(*
SPDX-FileCopyrightText: © 2026 Oleksandr Tiutyk <trofimich@gmail.com>
SPDX-License-Identifier: MIT
License: https://opensource.org/license/mit
*)

(*!
<summary>Verifies the testing library with an independent cyclic driver and direct expectations.</summary>
<description>
Runs sixteen scenarios in order with separate inner runners, including deliberately failed inner tests.
Keeps fixtures and the first diagnostic alive across scans. Publishes results directly to the ADS log.
Call Execute once per scan in the owning test task. AutomationRunner owns task memory cleanup.
This suite runs once per application initialization. Do not copy fixture state.
</description>
*)

{attribute 'no_assign'}
{attribute 'no_explicit_call' := 'do not call this function block directly'}
FUNCTION_BLOCK TestRunnerContractTest
VAR_STAT
	{attribute 'hide'}
	_ClassName : STRING := __POUNAME();
END_VAR
VAR CONSTANT
	//! <summary>Number of scenarios scheduled by the independent driver.</summary>
	_TestCount : DINT := 16;
	//! <summary>Maximum calls allowed for the empty runner to report completion.</summary>
	_EmptyScanLimit : UDINT := 16;
	//! <summary>Maximum calls per deadline phase on the configured 10 ms TestTask.</summary>
	_DeadlineScanLimit : UDINT := 32;
END_VAR
VAR_OUTPUT
	//! <summary>Number of completed scenarios with no outer assertion failures.</summary>
	PassedTests : DINT;
	//! <summary>Number of completed scenarios with an outer assertion failure or an unexpected exception.</summary>
	FailedTests : DINT;
	//! <summary>TRUE after every scenario has an outcome and the summary has been published.</summary>
	IsFinished : BOOL;
END_VAR
VAR
	_Scenario : TEST_RUNNER_CONTRACT_SCENARIO;
	_CaseFailed : BOOL;
	_FailureMessage : STRING(255);
END_VAR
VAR
	_Runner : MixedTestRunner;
	_Reporter : TOF_Testing.JUnitXmlReporter;
	_Configured : BOOL;
	_Calls : UDINT;
	_Repeated : BOOL;

	_FailingRun : IsolationTestRunner;
	_PassingRun : AssertionCallerTestRunner;
	_FailureReport : TOF_Testing.JUnitXmlReporter;
	_PassReport : TOF_Testing.JUnitXmlReporter;
	_IsolationConfigured : BOOL;
	_IsolationSecondRun : BOOL;
	_IsolationCalls : UDINT;

	_EmptyRun : EmptyTestRunner;
	_EmptyReport : TOF_Testing.JUnitXmlReporter;
	_EmptyConfigured : BOOL;
	_EmptyCalls : UDINT;
	_AbortRun : ReporterAbortTestRunner;
	_AbortReport : ThrowingTestReporter;
	_InvalidReport : TOF_Testing.JUnitXmlReporter;
	_AbortConfigured : BOOL;
	_AbortCalls : UDINT;
	_AbortPostCalls : UDINT;

	_DeadlineRun : DeadlineTestRunner;
	_DeadlineReport : TOF_Testing.JUnitXmlReporter;
	_DeadlineConfigured : BOOL;
	_DeadlineBusyFailureRun : BOOL;
	_DeadlineCalls : UDINT;
	_ActiveConfigurationChecked : BOOL;

	_DuplicateGroup : PairTestGroup(name := "Duplicates", parent := 0);
	_ParentGroup : SingleChildTestGroup(name := "Parent", parent := _ChildGroup);
	_ChildGroup : SingleChildTestGroup(name := "Child", parent := _ParentGroup);
	_IndexedGroup : PairTestGroup(name := "Indexed children", parent := 0);

	_AbortRecoveryReport : TOF_Testing.JUnitXmlReporter;
	_AbortRecovered : BOOL;
	_ExternalRun : ExternalRecoveryTestRunner;
	_ExternalReport : TOF_Testing.JUnitXmlReporter;
	_ExternalConfigured : BOOL;
	_ExternalRecovered : BOOL;
	_ExternalCalls : UDINT;

	_DiagnosticRun : DiagnosticTestRunner;
	_DiagnosticReport : TOF_Testing.JUnitXmlReporter;
	_DiagnosticConfigured : BOOL;
	_DiagnosticCalls : UDINT;

	_AssertionRun : AssertionTestRunner;
	_AssertionReport : TOF_Testing.JUnitXmlReporter;
	_AssertionsConfigured : BOOL;
	_AssertionCalls : UDINT;

	_XmlReport : TOF_Testing.JUnitXmlReporter;

	_RootTopologyRunner : RootTopologyTestRunner;
	_RootTopologyReport : TOF_Testing.JUnitXmlReporter;
	_RootTopologyConfigured : BOOL;
	_RootTopologyCalls : UDINT;

	_MissingConfigurationGroup : MissingChildrenTestGroup(name := "Missing configuration", parent := 0);
	_MissingConfigurationRunner : MissingChildrenTestRunner;
	_ExceptionAdsReporter : TOF_Testing.AdsLogReporter;
	_AdsSummaryReporter : CapturingAdsLogReporter;

	//! <summary>Synthetic Parent chains for path observation only; these fixtures are not executed as trees.</summary>
	_PathRoot : EmptyTestGroup(
		name := "AAAAAAAAAAAAAAAAAAAAAAAAAAAAAAAAAAAAAAAAAAAAAAAAAAAAAAAAAAAAAAAAAAAAAAAAAAAAAAAA",
		parent := 0
	);
	_PathSecond : EmptyTestGroup(
		name := "BBBBBBBBBBBBBBBBBBBBBBBBBBBBBBBBBBBBBBBBBBBBBBBBBBBBBBBBBBBBBBBBBBBBBBBBBBBBBBBB",
		parent := _PathRoot
	);
	_PathThird : EmptyTestGroup(
		name := "CCCCCCCCCCCCCCCCCCCCCCCCCCCCCCCCCCCCCCCCCCCCCCCCCCCCCCCCCCCCCCCCCCCCCCCCCCCCCCCC",
		parent := _PathSecond
	);
	_PathFourth : EmptyTestGroup(
		name := "DDDDDDDDDDDDDDDDDDDDDDDDDDDDDDDDDDDDDDDDDDDDDDDDDDDDDDDDDDDDDDDDDDDDDDDDDDDDDDDD",
		parent := _PathThird
	);
	_PathEmpty : EmptyTestGroup(name := "", parent := _PathRoot);
	_PathUnicode : TestingProbe(name := "Ω", parent := _PathEmpty);
	//! <summary>Supplies 81 characters to exercise ordinary truncation at the 80-character name input.</summary>
	_PathLongNameInput : WSTRING(81) := "AAAAAAAAAAAAAAAAAAAAAAAAAAAAAAAAAAAAAAAAAAAAAAAAAAAAAAAAAAAAAAAAAAAAAAAAAAAAAAAAB";
	_PathLongName : EmptyTestGroup(
		name := _PathLongNameInput,
		parent := 0
	);
	_ReportPathRoot : EmptyTestGroup(name := "Report root", parent := 0);
	_ReportPathMiddle : EmptyTestGroup(name := "Middle", parent := _ReportPathRoot);
	_ReportPathInner : EmptyTestGroup(name := "Inner", parent := _ReportPathMiddle);
	_PathReport : TOF_Testing.JUnitXmlReporter;
	_MetadataBoolAssertionContext : TOF_Testing.BoolAssertionContext;
	_MetadataByteAssertionContext : TOF_Testing.ByteAssertionContext;
	_MetadataDateAssertionContext : TOF_Testing.DateAssertionContext;
	_MetadataDateTimeAssertionContext : TOF_Testing.DateTimeAssertionContext;
	_MetadataDIntAssertionContext : TOF_Testing.DIntAssertionContext;
	_MetadataDWordAssertionContext : TOF_Testing.DWordAssertionContext;
	_MetadataIntAssertionContext : TOF_Testing.IntAssertionContext;
	_MetadataLIntAssertionContext : TOF_Testing.LIntAssertionContext;
	_MetadataLongDateAssertionContext : TOF_Testing.LongDateAssertionContext;
	_MetadataLongDateTimeAssertionContext : TOF_Testing.LongDateTimeAssertionContext;
	_MetadataLongRealAssertionContext : TOF_Testing.LongRealAssertionContext;
	_MetadataLongTimeAssertionContext : TOF_Testing.LongTimeAssertionContext;
	_MetadataLongTimeOfDayAssertionContext : TOF_Testing.LongTimeOfDayAssertionContext;
	_MetadataLWordAssertionContext : TOF_Testing.LWordAssertionContext;
	_MetadataPointerAssertionContext : TOF_Testing.PointerAssertionContext;
	_MetadataRealAssertionContext : TOF_Testing.RealAssertionContext;
	_MetadataSIntAssertionContext : TOF_Testing.SIntAssertionContext;
	_MetadataStringAssertionContext : TOF_Testing.StringAssertionContext;
	_MetadataTimeAssertionContext : TOF_Testing.TimeAssertionContext;
	_MetadataTimeOfDayAssertionContext : TOF_Testing.TimeOfDayAssertionContext;
	_MetadataUDIntAssertionContext : TOF_Testing.UDIntAssertionContext;
	_MetadataUIntAssertionContext : TOF_Testing.UIntAssertionContext;
	_MetadataULIntAssertionContext : TOF_Testing.ULIntAssertionContext;
	_MetadataUSIntAssertionContext : TOF_Testing.USIntAssertionContext;
	_MetadataWideStringAssertionContext : TOF_Testing.WideStringAssertionContext;
	_MetadataWordAssertionContext : TOF_Testing.WordAssertionContext;
	_OtherBoolContext : TOF_Testing.BoolAssertionContext;
END_VAR

(*!
<summary>Advances one scenario and reports its outcome after completion.</summary>
<description>
Retains the first failed expectation across pending cycles. An unexpected exception fails the active scenario.
Checks the allocation latch outside the recovery block. The caller owns task memory cleanup.
Returns immediately after all scenarios finish and publishes exactly one summary per initialization.
</description>
*)
METHOD Execute
VAR
	caseName : STRING(80);
	nextScenario : TEST_RUNNER_CONTRACT_SCENARIO;
	completed : BOOL;
	exceptionCode : __SYSTEM.ExceptionCode;
END_VAR
IF IsFinished THEN
	RETURN;
END_IF

IF _Scenario = TEST_RUNNER_CONTRACT_SCENARIO.STARTING THEN
	logResult(isError := FALSE, message := TOF_Core.Strings.Concat255('Starting ', TO_STRING(_TestCount), ' tests'));
	_Scenario := TEST_RUNNER_CONTRACT_SCENARIO.ELEMENT_TREE;

	RETURN;
END_IF

__TRY
	CASE _Scenario OF
		TEST_RUNNER_CONTRACT_SCENARIO.ELEMENT_TREE:
			caseName := 'Element tree, lifecycle, repeated run and JUnit';
			nextScenario := TEST_RUNNER_CONTRACT_SCENARIO.CASE_ISOLATION;
			completed := runAndCheck();

		TEST_RUNNER_CONTRACT_SCENARIO.CASE_ISOLATION:
			caseName := 'Each failure belongs to its receiving case';
			nextScenario := TEST_RUNNER_CONTRACT_SCENARIO.EMPTY_RUN;
			completed := checkCaseIsolation();

		TEST_RUNNER_CONTRACT_SCENARIO.EMPTY_RUN:
			caseName := 'An empty root passes with zero tests';
			nextScenario := TEST_RUNNER_CONTRACT_SCENARIO.REPORTER_ABORT;
			completed := checkEmptyRun();

		TEST_RUNNER_CONTRACT_SCENARIO.REPORTER_ABORT:
			caseName := 'A throwing reporter aborts without retry';
			nextScenario := TEST_RUNNER_CONTRACT_SCENARIO.DEADLINE;
			completed := checkReporterAbort();

		TEST_RUNNER_CONTRACT_SCENARIO.DEADLINE:
			caseName := 'A pending multi-cycle test fails at its deadline';
			nextScenario := TEST_RUNNER_CONTRACT_SCENARIO.GROUP_TOPOLOGY;
			completed := checkDeadline();

		TEST_RUNNER_CONTRACT_SCENARIO.GROUP_TOPOLOGY:
			caseName := 'Static group topology is validated before child callbacks';
			nextScenario := TEST_RUNNER_CONTRACT_SCENARIO.EXTERNAL_RECOVERY;
			completed := checkTopology();

		TEST_RUNNER_CONTRACT_SCENARIO.EXTERNAL_RECOVERY:
			caseName := 'External abort recovery can be retried for the same static tree';
			nextScenario := TEST_RUNNER_CONTRACT_SCENARIO.DIAGNOSTICS;
			completed := checkExternalRecovery();

		TEST_RUNNER_CONTRACT_SCENARIO.DIAGNOSTICS:
			caseName := 'Native and framework diagnostics outlive their exception objects';
			nextScenario := TEST_RUNNER_CONTRACT_SCENARIO.ADS_REPORTER_SUMMARY;
			completed := checkDiagnostics();

		TEST_RUNNER_CONTRACT_SCENARIO.ADS_REPORTER_SUMMARY:
			caseName := 'ADS summary retains first failure and resets on the next run';
			nextScenario := TEST_RUNNER_CONTRACT_SCENARIO.ASSERTION_CONTRACTS;
			completed := checkAdsReporterSummary();

		TEST_RUNNER_CONTRACT_SCENARIO.ASSERTION_CONTRACTS:
			caseName := 'Independent contexts, typed predicates, snapshots and chain diagnostics';
			nextScenario := TEST_RUNNER_CONTRACT_SCENARIO.XML_ENCODING;
			completed := checkAssertionContracts();

		TEST_RUNNER_CONTRACT_SCENARIO.XML_ENCODING:
			caseName := 'JUnit preserves long text and replaces forbidden Unicode sequences';
			nextScenario := TEST_RUNNER_CONTRACT_SCENARIO.RUNNER_TOPOLOGY;
			completed := checkXmlEncoding();

		TEST_RUNNER_CONTRACT_SCENARIO.RUNNER_TOPOLOGY:
			caseName := 'Static runner validates roots at startup and executes without rescanning';
			nextScenario := TEST_RUNNER_CONTRACT_SCENARIO.EXCEPTION_CLASSES;
			completed := checkRunnerTopology();

		TEST_RUNNER_CONTRACT_SCENARIO.EXCEPTION_CLASSES:
			caseName := 'Missing static storage is diagnosed before child access';
			nextScenario := TEST_RUNNER_CONTRACT_SCENARIO.CONTEXT_OBJECTS;
			completed := checkExceptionClasses();

		TEST_RUNNER_CONTRACT_SCENARIO.CONTEXT_OBJECTS:
			caseName := 'Typed contexts and concrete runner expose Object metadata and identity';
			nextScenario := TEST_RUNNER_CONTRACT_SCENARIO.PATHS;
			completed := checkContextObjects();

		TEST_RUNNER_CONTRACT_SCENARIO.PATHS:
			caseName := 'Paths follow live Parent links without Reset context';
			nextScenario := TEST_RUNNER_CONTRACT_SCENARIO.INDEXED_CHILDREN;
			completed := checkPaths();

		TEST_RUNNER_CONTRACT_SCENARIO.INDEXED_CHILDREN:
			caseName := 'Indexed children preserve order and reject missing storage or invalid indices';
			nextScenario := TEST_RUNNER_CONTRACT_SCENARIO.FINISHED;
			completed := checkIndexedChildren();
	ELSE
		caseName := 'Scenario selection';
		nextScenario := TEST_RUNNER_CONTRACT_SCENARIO.FINISHED;
		expect(condition := FALSE, message := 'Invalid scenario selection');
		completed := TRUE;
	END_CASE
__CATCH(exceptionCode)
	expect(
		condition := FALSE,
		message := TOF_Core.Strings.Concat255('Unexpected PLC exception ', TO_STRING(exceptionCode))
	);
	completed := TRUE;
__ENDTRY

TOF_Core.DynamicMemoryManager.RaiseIfAllocationFailed();

IF NOT completed THEN
	RETURN;
END_IF

IF _CaseFailed THEN
	FailedTests := FailedTests + 1;
	logResult(
		isError := TRUE,
		message := TOF_Core.Strings.Concat255(caseName, ': ', _FailureMessage)
	);
ELSE
	PassedTests := PassedTests + 1;
END_IF

_CaseFailed := FALSE;
_FailureMessage := '';
_Scenario := nextScenario;

IF _Scenario = TEST_RUNNER_CONTRACT_SCENARIO.FINISHED THEN
	logResult(
		isError := FailedTests <> 0,
		message := TOF_Core.Strings.Concat255(
			'Finished: ',
			TO_STRING(PassedTests),
			' passed, ',
			TO_STRING(FailedTests),
			' failed'
		)
	);
	IsFinished := TRUE;
END_IF
END_METHOD

(*!
<summary>Copies the first diagnostic when an expectation fails.</summary>
<param name="condition">TRUE when the expectation holds.</param>
<param name="message">Description of the failed expectation.</param>
*)
METHOD PRIVATE expect
VAR_INPUT
	condition : BOOL;
	message : STRING(255);
END_VAR
IF NOT condition AND_THEN NOT _CaseFailed THEN
	_CaseFailed := TRUE;
	_FailureMessage := message;
END_IF
END_METHOD

(*!
<summary>Checks that a predicate is false.</summary>
<param name="condition">Predicate that must be FALSE.</param>
<param name="message">Description of the failed expectation.</param>
*)
METHOD PRIVATE expectFalse
VAR_INPUT
	condition : BOOL;
	message : STRING(255);
END_VAR
expect(condition := NOT condition, message := message);
END_METHOD

(*!
<summary>Compares two DINT values and records differences.</summary>
<param name="expected">Expected value determined by the scenario.</param>
<param name="actual">Observed value.</param>
<param name="message">Description of the failed expectation.</param>
*)
METHOD PRIVATE expectDInt
VAR_INPUT
	expected : DINT;
	actual : DINT;
	message : STRING(255);
END_VAR
IF actual <> expected AND_THEN NOT _CaseFailed THEN
	expect(
		condition := FALSE,
		message := TOF_Core.Strings.Concat255(
			message,
			' (expected ',
			TO_STRING(expected),
			', actual ',
			TO_STRING(actual),
			')'
		)
	);
END_IF
END_METHOD

(*!
<summary>Compares two UDINT values and records differences.</summary>
<param name="expected">Expected value determined by the scenario.</param>
<param name="actual">Observed value.</param>
<param name="message">Description of the failed expectation.</param>
*)
METHOD PRIVATE expectUDInt
VAR_INPUT
	expected : UDINT;
	actual : UDINT;
	message : STRING(255);
END_VAR
IF actual <> expected AND_THEN NOT _CaseFailed THEN
	expect(
		condition := FALSE,
		message := TOF_Core.Strings.Concat255(
			message,
			' (expected ',
			TO_STRING(expected),
			', actual ',
			TO_STRING(actual),
			')'
		)
	);
END_IF
END_METHOD

(*!
<summary>Publishes a diagnostic without using the library under test.</summary>
<param name="isError">TRUE for scenario errors and failed summaries.</param>
<param name="message">Diagnostic to publish.</param>
*)
METHOD PRIVATE logResult
VAR_INPUT
	isError : BOOL;
	message : STRING(255);
END_VAR
VAR
	severity : DWORD;
END_VAR
severity := SEL(
	isError,
	Tc2_System.Global_Variables.ADSLOG_MSGTYPE_HINT,
	Tc2_System.Global_Variables.ADSLOG_MSGTYPE_ERROR
);

Tc2_System.ADSLOGSTR(
	msgCtrlMask := severity OR Tc2_System.Global_Variables.ADSLOG_MSGTYPE_LOG,
	msgFmtStr := '[TestRunnerContractTest] %s',
	strArg := message
);
END_METHOD

(*!
<summary>Checks a caught failure through its dedicated exception interface before task cleanup.</summary>
<description>Only borrows the exception during this call; no exception reference survives the test cycle.</description>
*)
METHOD PRIVATE assertCaughtExceptionType
VAR_INPUT
	exceptionCode : __SYSTEM.ExceptionCode;
	expectedTypeName : STRING;
END_VAR
VAR
	exception : TOF_Core.IException;
	standardException : TOF_Core.IStandardException;
	argumentNotSpecified : TOF_Core.IArgumentNotSpecifiedException;
	memberNotSpecified : TOF_Core.IDataMemberNotSpecifiedException;
	argumentValueNotSupported : TOF_Core.IArgumentValueNotSupportedException;
	argumentOutOfRange : TOF_Core.IArgumentOutOfRangeException;
	matchesType : BOOL;
END_VAR
exception := TOF_Core.ExceptionManager.GetLastException(
	exceptionCode := exceptionCode,
	catchPointNamespaceName := CurrentNamespace.Name,
	catchPointPOUName := __POUNAME(),
	catchPointPosition := __POSITION()
);
expect(condition := exception <> 0, message := 'Caught failure exposes its exception payload');

IF exception = 0 THEN
	RETURN;
END_IF

IF expectedTypeName = 'StandardException' THEN
	matchesType := __QUERYINTERFACE(exception, standardException);
ELSIF expectedTypeName = 'ArgumentNotSpecifiedException' THEN
	matchesType := __QUERYINTERFACE(exception, argumentNotSpecified);
ELSIF expectedTypeName = 'DataMemberNotSpecifiedException' THEN
	matchesType := __QUERYINTERFACE(exception, memberNotSpecified);
ELSIF expectedTypeName = 'ArgumentValueNotSupportedException' THEN
	matchesType := __QUERYINTERFACE(exception, argumentValueNotSupported);
ELSIF expectedTypeName = 'ArgumentOutOfRangeException' THEN
	matchesType := __QUERYINTERFACE(exception, argumentOutOfRange);
END_IF

expect(condition := matchesType, message := 'Exception interface matches the expected failure category');
END_METHOD

(*!
<summary>Checks concrete metadata through a borrowed Object interface.</summary>
<description>Checks namespace, class, size and address separately with distinct failure diagnostics.</description>
<param name="object">Live instance whose metadata is read without preparation.</param>
<param name="expectedNamespaceName">Namespace of the project declaring the concrete type.</param>
<param name="expectedClassName">Concrete context class name.</param>
<param name="expectedSize">Compiler-reported size of the complete concrete context.</param>
<param name="expectedAddress">Address of the concrete context, without ownership transfer.</param>
*)
METHOD PRIVATE assertObjectMetadata
VAR_INPUT
	object : TOF_Core.IObject;
	expectedNamespaceName : STRING;
	expectedClassName : STRING;
	expectedSize : ULINT;
	expectedAddress : PVOID;
END_VAR
expect(condition := object <> 0, message := expectedClassName);

IF object = 0 THEN
	RETURN;
END_IF

expect(
	condition := object.ClassName = expectedClassName,
	message := TOF_Core.Strings.Concat255(expectedClassName, ': ClassName')
);
expect(
	condition := object.NamespaceName = expectedNamespaceName,
	message := TOF_Core.Strings.Concat255(expectedClassName, ': NamespaceName')
);
expect(
	condition := object.SelfSize = expectedSize,
	message := TOF_Core.Strings.Concat255(expectedClassName, ': SelfSize')
);
expect(
	condition := object.SelfAddress = expectedAddress,
	message := TOF_Core.Strings.Concat255(expectedClassName, ': SelfAddress')
);
END_METHOD

(*!
<summary>Checks independent typed and generic contexts, native predicates and chain-wide diagnostics.</summary>
<description>Configures the persistent output probes through a local reference without copying them.
Returns TRUE when all observations for this scenario are complete.
</description>
*)
METHOD PRIVATE checkAssertionContracts : BOOL
VAR
	probe : REFERENCE TO AssertionContractProbe;
END_VAR
IF NOT _AssertionsConfigured THEN
	probe REF= _AssertionRun.Assertion0;
	probe.Scenario := ASSERTION_PROBE_SCENARIO.FLOAT_TOLERANCE;
	probe REF= _AssertionRun.Assertion1;
	probe.Scenario := ASSERTION_PROBE_SCENARIO.INTEGER_EXACT;
	probe REF= _AssertionRun.Assertion2;
	probe.Scenario := ASSERTION_PROBE_SCENARIO.TYPED_LITERALS;
	probe REF= _AssertionRun.Assertion3;
	probe.Scenario := ASSERTION_PROBE_SCENARIO.MESSAGE_CHAIN;
	probe REF= _AssertionRun.Assertion4;
	probe.Scenario := ASSERTION_PROBE_SCENARIO.NEGATIVE_TOLERANCE;
	probe REF= _AssertionRun.Assertion5;
	probe.Scenario := ASSERTION_PROBE_SCENARIO.NAN_TOLERANCE;
	probe REF= _AssertionRun.Assertion6;
	probe.Scenario := ASSERTION_PROBE_SCENARIO.INFINITE_TOLERANCE;
	probe REF= _AssertionRun.Assertion7;
	probe.Scenario := ASSERTION_PROBE_SCENARIO.MESSAGE_RESET;
	probe REF= _AssertionRun.Assertion8;
	probe.Scenario := ASSERTION_PROBE_SCENARIO.POINTERS_AND_STRINGS;
	probe REF= _AssertionRun.Assertion9;
	probe.Scenario := ASSERTION_PROBE_SCENARIO.FIRST_FAILURE;
	probe REF= _AssertionRun.Assertion10;
	probe.Scenario := ASSERTION_PROBE_SCENARIO.SPECIAL_FLOATS;
	probe REF= _AssertionRun.Assertion11;
	probe.Scenario := ASSERTION_PROBE_SCENARIO.OPPOSITE_LIMITS;
	probe REF= _AssertionRun.Assertion12;
	probe.Scenario := ASSERTION_PROBE_SCENARIO.GENERIC_MESSAGE_CHAIN;
	probe REF= _AssertionRun.Assertion13;
	probe.Scenario := ASSERTION_PROBE_SCENARIO.GENERIC_MESSAGE_RESET;
	probe REF= _AssertionRun.Assertion14;
	probe.Scenario := ASSERTION_PROBE_SCENARIO.CONTEXT_TRANSITIONS;
	probe REF= _AssertionRun.Assertion15;
	probe.Scenario := ASSERTION_PROBE_SCENARIO.TYPED_MESSAGE_AFTER_GENERIC;
	probe REF= _AssertionRun.Assertion16;
	probe.Scenario := ASSERTION_PROBE_SCENARIO.GENERIC_MESSAGE_AFTER_TYPED;
	probe REF= _AssertionRun.Assertion17;
	probe.Scenario := ASSERTION_PROBE_SCENARIO.TYPED_MESSAGE_RESET_AFTER_GENERIC;
	probe REF= _AssertionRun.Assertion18;
	probe.Scenario := ASSERTION_PROBE_SCENARIO.INTEGER_FAILURE;
	probe REF= _AssertionRun.Assertion19;
	probe.Scenario := ASSERTION_PROBE_SCENARIO.BITSTRING_FAILURE;
	probe REF= _AssertionRun.Assertion20;
	probe.Scenario := ASSERTION_PROBE_SCENARIO.POINTER_FAILURE;
	probe REF= _AssertionRun.Assertion21;
	probe.Scenario := ASSERTION_PROBE_SCENARIO.STRING_LONG_FAILURE;
	probe REF= _AssertionRun.Assertion22;
	probe.Scenario := ASSERTION_PROBE_SCENARIO.WIDE_STRING_LONG_FAILURE;
	probe REF= _AssertionRun.Assertion23;
	probe.Scenario := ASSERTION_PROBE_SCENARIO.STRING_CONTAINMENT_FAILURE;
	probe REF= _AssertionRun.Assertion24;
	probe.Scenario := ASSERTION_PROBE_SCENARIO.FLOAT_ORDERING_FAILURE;
	probe REF= _AssertionRun.Assertion25;
	probe.Scenario := ASSERTION_PROBE_SCENARIO.FLOAT_EQUALITY_FAILURE;
	probe REF= _AssertionRun.Assertion26;
	probe.Scenario := ASSERTION_PROBE_SCENARIO.TIME_ORDERING_FAILURE;
	_AssertionRun.Reporter := _AssertionReport;
	_AssertionsConfigured := TRUE;
END_IF

_AssertionRun.Execute(cleanupTaskMemory := FALSE);
_AssertionCalls := _AssertionCalls + 1;

IF NOT _AssertionRun.IsFinished AND_THEN _AssertionCalls < 32 THEN
	RETURN;
END_IF

expect(condition := _AssertionRun.IsFinished, message := 'Twenty-seven assertion leaves finish within 32 scans');
expectDInt(expected := 27, actual := _AssertionRun.TotalTests, message := 'Every assertion scenario executes');
expectDInt(
	expected := 7,
	actual := _AssertionRun.PassedTests,
	message := 'Seven supported assertion scenarios pass'
);
expectDInt(
	expected := 20,
	actual := _AssertionRun.FailedTests,
	message := 'Twenty deliberate failures are recorded'
);
expect(
	condition := _AssertionRun.Assertion0.Outcome = TOF_Testing.TEST_OUTCOME.PASSED,
	message := 'Assertion scenario 0 has its expected passed outcome'
);
expect(
	condition := _AssertionRun.Assertion1.Outcome = TOF_Testing.TEST_OUTCOME.PASSED,
	message := 'Assertion scenario 1 has its expected passed outcome'
);
expect(
	condition := _AssertionRun.Assertion2.Outcome = TOF_Testing.TEST_OUTCOME.PASSED,
	message := 'Assertion scenario 2 has its expected passed outcome'
);
expect(
	condition := _AssertionRun.Assertion3.Outcome = TOF_Testing.TEST_OUTCOME.FAILED,
	message := 'Assertion scenario 3 has its expected failed outcome'
);
expect(
	condition := _AssertionRun.Assertion4.Outcome = TOF_Testing.TEST_OUTCOME.FAILED,
	message := 'Assertion scenario 4 has its expected failed outcome'
);
expect(
	condition := _AssertionRun.Assertion5.Outcome = TOF_Testing.TEST_OUTCOME.FAILED,
	message := 'Assertion scenario 5 has its expected failed outcome'
);
expect(
	condition := _AssertionRun.Assertion6.Outcome = TOF_Testing.TEST_OUTCOME.FAILED,
	message := 'Assertion scenario 6 has its expected failed outcome'
);
expect(
	condition := _AssertionRun.Assertion7.Outcome = TOF_Testing.TEST_OUTCOME.FAILED,
	message := 'Assertion scenario 7 has its expected failed outcome'
);
expect(
	condition := _AssertionRun.Assertion8.Outcome = TOF_Testing.TEST_OUTCOME.PASSED,
	message := 'Assertion scenario 8 has its expected passed outcome'
);
expect(
	condition := _AssertionRun.Assertion9.Outcome = TOF_Testing.TEST_OUTCOME.FAILED,
	message := 'Assertion scenario 9 has its expected failed outcome'
);
expect(
	condition := _AssertionRun.Assertion10.Outcome = TOF_Testing.TEST_OUTCOME.PASSED,
	message := 'Assertion scenario 10 has its expected passed outcome'
);
expect(
	condition := _AssertionRun.Assertion11.Outcome = TOF_Testing.TEST_OUTCOME.PASSED,
	message := 'Assertion scenario 11 has its expected passed outcome'
);
expect(
	condition := _AssertionRun.Assertion12.Outcome = TOF_Testing.TEST_OUTCOME.FAILED,
	message := 'Assertion scenario 12 has its expected failed outcome'
);
expect(
	condition := _AssertionRun.Assertion13.Outcome = TOF_Testing.TEST_OUTCOME.FAILED,
	message := 'Assertion scenario 13 has its expected failed outcome'
);
expect(
	condition := _AssertionRun.Assertion9.FailureMessage = "First diagnostic",
	message := 'Later assertion and teardown exception preserve the first failure'
);
expect(
	condition := TOF_Core.WideStrings.Contains(
		stringToSearchIn := _AssertionRun.Assertion3.FailureMessage,
		stringToFind := "Chain diagnostic: Expected value < "
	),
	message := 'The message survives a successful assertion in the same typed chain'
);
expect(
	condition := NOT TOF_Core.WideStrings.Contains(
		stringToSearchIn := _AssertionRun.Assertion7.FailureMessage,
		stringToFind := "Previous diagnostic"
	),
	message := 'Omitting the typed entry message clears the previous prefix'
);
expect(
	condition := TOF_Core.WideStrings.Contains(
		stringToSearchIn := _AssertionRun.Assertion12.FailureMessage,
		stringToFind := "Generic chain diagnostic: Expected value < "
	),
	message := 'Borrowed assertions retain the same chain-wide message contract'
);
expect(
	condition := NOT TOF_Core.WideStrings.Contains(
		stringToSearchIn := _AssertionRun.Assertion13.FailureMessage,
		stringToFind := "Previous generic diagnostic"
	),
	message := 'Omitting the borrowed entry message clears the previous prefix'
);
expect(
	condition := TOF_Core.WideStrings.Contains(
		stringToSearchIn := _AssertionRun.Assertion4.FailureMessage,
		stringToFind := "finite nonnegative comparison tolerance"
	),
	message := 'An invalid tolerance fails before a comparison that would otherwise pass'
);
expect(
	condition := _AssertionRun.Assertion14.Outcome = TOF_Testing.TEST_OUTCOME.PASSED,
	message := 'Independent context scenario CONTEXT_TRANSITIONS has its expected outcome'
);
expect(
	condition := _AssertionRun.Assertion15.Outcome = TOF_Testing.TEST_OUTCOME.FAILED,
	message := 'Independent context scenario TYPED_MESSAGE_AFTER_GENERIC has its expected outcome'
);
expect(
	condition := _AssertionRun.Assertion15.FailureMessage = "Independent typed: Expected: 11, but was: 10",
	message := 'Independent context scenario TYPED_MESSAGE_AFTER_GENERIC retains its diagnostic'
);
expect(
	condition := _AssertionRun.Assertion16.Outcome = TOF_Testing.TEST_OUTCOME.FAILED,
	message := 'Independent context scenario GENERIC_MESSAGE_AFTER_TYPED has its expected outcome'
);
expect(
	condition := _AssertionRun.Assertion16.FailureMessage = "Independent generic: Expected: 2, but was: 1",
	message := 'Independent context scenario GENERIC_MESSAGE_AFTER_TYPED retains its diagnostic'
);
expect(
	condition := _AssertionRun.Assertion17.Outcome = TOF_Testing.TEST_OUTCOME.FAILED,
	message := 'Independent context scenario TYPED_MESSAGE_RESET_AFTER_GENERIC has its expected outcome'
);
expect(
	condition := _AssertionRun.Assertion17.FailureMessage = "Expected: 2, but was: 1",
	message := 'Independent context scenario TYPED_MESSAGE_RESET_AFTER_GENERIC retains its diagnostic'
);
expect(
	condition := _AssertionRun.Assertion18.Outcome = TOF_Testing.TEST_OUTCOME.FAILED,
	message := 'Independent context scenario INTEGER_FAILURE has its expected outcome'
);
expect(
	condition := _AssertionRun.Assertion18.FailureMessage = "Expected: -2, but was: -3",
	message := 'Independent context scenario INTEGER_FAILURE retains its diagnostic'
);
expect(
	condition := _AssertionRun.Assertion19.Outcome = TOF_Testing.TEST_OUTCOME.FAILED,
	message := 'Independent context scenario BITSTRING_FAILURE has its expected outcome'
);
expect(
	condition := _AssertionRun.Assertion19.FailureMessage = "Expected: 11, but was: 10",
	message := 'Independent context scenario BITSTRING_FAILURE retains its diagnostic'
);
expect(
	condition := _AssertionRun.Assertion20.Outcome = TOF_Testing.TEST_OUTCOME.FAILED,
	message := 'Independent context scenario POINTER_FAILURE has its expected outcome'
);
expect(
	condition := TOF_Core.WideStrings.Contains(
		stringToSearchIn := _AssertionRun.Assertion20.FailureMessage,
		stringToFind := "Expected: 0, but was: "
	),
	message := 'Independent context scenario POINTER_FAILURE retains its diagnostic'
);
expect(
	condition := _AssertionRun.Assertion21.Outcome = TOF_Testing.TEST_OUTCOME.FAILED,
	message := 'Independent context scenario STRING_LONG_FAILURE has its expected outcome'
);
expect(
	condition := TOF_Core.WideStrings.Contains(
		stringToSearchIn := _AssertionRun.Assertion21.FailureMessage,
		stringToFind := "ASCII expected suffix"
	),
	message := 'Independent context scenario STRING_LONG_FAILURE retains its diagnostic'
);
expect(
	condition := _AssertionRun.Assertion22.Outcome = TOF_Testing.TEST_OUTCOME.FAILED,
	message := 'Independent context scenario WIDE_STRING_LONG_FAILURE has its expected outcome'
);
expect(
	condition := TOF_Core.WideStrings.Contains(
		stringToSearchIn := _AssertionRun.Assertion22.FailureMessage,
		stringToFind := "Wide expected suffix"
	),
	message := 'Independent context scenario WIDE_STRING_LONG_FAILURE retains its diagnostic'
);
expect(
	condition := _AssertionRun.Assertion23.Outcome = TOF_Testing.TEST_OUTCOME.FAILED,
	message := 'Independent context scenario STRING_CONTAINMENT_FAILURE has its expected outcome'
);
expect(
	condition := _AssertionRun.Assertion23.FailureMessage = "Expected text to contain 'missing', but was: 'present'",
	message := 'Independent context scenario STRING_CONTAINMENT_FAILURE retains its diagnostic'
);
expect(
	condition := _AssertionRun.Assertion24.Outcome = TOF_Testing.TEST_OUTCOME.FAILED,
	message := 'Independent context scenario FLOAT_ORDERING_FAILURE has its expected outcome'
);
expect(
	condition := TOF_Core.WideStrings.Contains(
		stringToSearchIn := _AssertionRun.Assertion24.FailureMessage,
		stringToFind := "Expected value > "
	),
	message := 'Independent context scenario FLOAT_ORDERING_FAILURE retains its diagnostic'
);
expect(
	condition := _AssertionRun.Assertion25.Outcome = TOF_Testing.TEST_OUTCOME.FAILED,
	message := 'Independent context scenario FLOAT_EQUALITY_FAILURE has its expected outcome'
);
expect(
	condition := TOF_Core.WideStrings.Contains(
		stringToSearchIn := _AssertionRun.Assertion25.FailureMessage,
		stringToFind := ", tolerance: "
	),
	message := 'Independent context scenario FLOAT_EQUALITY_FAILURE retains its diagnostic'
);
expect(
	condition := _AssertionRun.Assertion26.Outcome = TOF_Testing.TEST_OUTCOME.FAILED,
	message := 'Independent context scenario TIME_ORDERING_FAILURE has its expected outcome'
);
expect(
	condition := TOF_Core.WideStrings.Contains(
		stringToSearchIn := _AssertionRun.Assertion26.FailureMessage,
		stringToFind := "Expected value >= "
	),
	message := 'Independent context scenario TIME_ORDERING_FAILURE retains its diagnostic'
);
checkAssertionContracts := TRUE;
END_METHOD

(*!
<summary>Checks assertion and direct failure routing between independent active cases.</summary>
<description>Configures the persistent output probes through local references without copying them.
Returns TRUE when all observations for this scenario are complete.
</description>
*)
METHOD PRIVATE checkCaseIsolation : BOOL
VAR
	passingProbe : REFERENCE TO AssertionIsolationProbe;
	failingProbe : REFERENCE TO AssertionIsolationProbe;
END_VAR
passingProbe REF= _PassingRun.Child;
failingProbe REF= _FailingRun.Child;

IF NOT _IsolationConfigured THEN
	passingProbe.Peer := ADR(failingProbe);
	failingProbe.Timeout := T#0S;
	passingProbe.Timeout := T#0S;
	_FailingRun.Reporter := _FailureReport;
	_PassingRun.Reporter := _PassReport;
	_IsolationConfigured := TRUE;
END_IF

_FailingRun.Execute(cleanupTaskMemory := FALSE);
_PassingRun.Execute(cleanupTaskMemory := FALSE);
_IsolationCalls := _IsolationCalls + 1;

IF NOT (_FailingRun.IsFinished AND_THEN _PassingRun.IsFinished) AND_THEN _IsolationCalls < 16 THEN
	RETURN;
END_IF

expect(condition := _FailingRun.IsFinished AND _PassingRun.IsFinished, message := 'Both runs finish');
expectDInt(expected := 1, actual := _FailingRun.FailedTests, message := 'Failure belongs to receiver');
expectDInt(expected := 1, actual := _PassingRun.PassedTests, message := 'Calling case passes');
expectDInt(expected := 0, actual := _PassingRun.FailedTests, message := 'Calling case has no peer failure');

IF NOT _IsolationSecondRun AND_THEN _FailingRun.IsFinished AND_THEN _PassingRun.IsFinished THEN
	_IsolationSecondRun := TRUE;
	passingProbe.UseDirectFailure := TRUE;
	_IsolationCalls := 0;
	_FailingRun.Reset();
	_PassingRun.Reset();
	RETURN;
END_IF

checkCaseIsolation := TRUE;
END_METHOD

(*!
<summary>Checks all typed contexts through IObject before assertion preparation.</summary>
<description>
Persistent contexts retain their default state. Checks metadata, addresses and inherited identity equality;
no test callback or Prepare call is required to read Object metadata.
Also checks concrete runner metadata, the inherited INamed signature and the constructor-copied group name.
Context namespaces are compared with an independent library reporter; runner metadata uses the consumer namespace.

Returns TRUE when all observations for this scenario are complete.
</description>
*)
METHOD PRIVATE checkContextObjects : BOOL
VAR
	first : TOF_Core.IObject;
	second : TOF_Core.IObject;
	group : TOF_Core.IObject;
	named : TOF_Core.INamed;
	displayName : REFERENCE TO WSTRING;
	concreteDisplayName : REFERENCE TO WSTRING;
END_VAR
assertObjectMetadata(
	object := _Runner,
	expectedNamespaceName := CurrentNamespace.Name,
	expectedClassName := 'MixedTestRunner',
	expectedSize := XSIZEOF(_Runner),
	expectedAddress := ADR(_Runner)
);

assertObjectMetadata(
	object := _MetadataBoolAssertionContext,
	expectedNamespaceName := _ExceptionAdsReporter.NamespaceName,
	expectedClassName := 'BoolAssertionContext',
	expectedSize := XSIZEOF(_MetadataBoolAssertionContext),
	expectedAddress := ADR(_MetadataBoolAssertionContext)
);
assertObjectMetadata(
	object := _MetadataByteAssertionContext,
	expectedNamespaceName := _ExceptionAdsReporter.NamespaceName,
	expectedClassName := 'ByteAssertionContext',
	expectedSize := XSIZEOF(_MetadataByteAssertionContext),
	expectedAddress := ADR(_MetadataByteAssertionContext)
);
assertObjectMetadata(
	object := _MetadataDateAssertionContext,
	expectedNamespaceName := _ExceptionAdsReporter.NamespaceName,
	expectedClassName := 'DateAssertionContext',
	expectedSize := XSIZEOF(_MetadataDateAssertionContext),
	expectedAddress := ADR(_MetadataDateAssertionContext)
);
assertObjectMetadata(
	object := _MetadataDateTimeAssertionContext,
	expectedNamespaceName := _ExceptionAdsReporter.NamespaceName,
	expectedClassName := 'DateTimeAssertionContext',
	expectedSize := XSIZEOF(_MetadataDateTimeAssertionContext),
	expectedAddress := ADR(_MetadataDateTimeAssertionContext)
);
assertObjectMetadata(
	object := _MetadataDIntAssertionContext,
	expectedNamespaceName := _ExceptionAdsReporter.NamespaceName,
	expectedClassName := 'DIntAssertionContext',
	expectedSize := XSIZEOF(_MetadataDIntAssertionContext),
	expectedAddress := ADR(_MetadataDIntAssertionContext)
);
assertObjectMetadata(
	object := _MetadataDWordAssertionContext,
	expectedNamespaceName := _ExceptionAdsReporter.NamespaceName,
	expectedClassName := 'DWordAssertionContext',
	expectedSize := XSIZEOF(_MetadataDWordAssertionContext),
	expectedAddress := ADR(_MetadataDWordAssertionContext)
);
assertObjectMetadata(
	object := _MetadataIntAssertionContext,
	expectedNamespaceName := _ExceptionAdsReporter.NamespaceName,
	expectedClassName := 'IntAssertionContext',
	expectedSize := XSIZEOF(_MetadataIntAssertionContext),
	expectedAddress := ADR(_MetadataIntAssertionContext)
);
assertObjectMetadata(
	object := _MetadataLIntAssertionContext,
	expectedNamespaceName := _ExceptionAdsReporter.NamespaceName,
	expectedClassName := 'LIntAssertionContext',
	expectedSize := XSIZEOF(_MetadataLIntAssertionContext),
	expectedAddress := ADR(_MetadataLIntAssertionContext)
);
assertObjectMetadata(
	object := _MetadataLongDateAssertionContext,
	expectedNamespaceName := _ExceptionAdsReporter.NamespaceName,
	expectedClassName := 'LongDateAssertionContext',
	expectedSize := XSIZEOF(_MetadataLongDateAssertionContext),
	expectedAddress := ADR(_MetadataLongDateAssertionContext)
);
assertObjectMetadata(
	object := _MetadataLongDateTimeAssertionContext,
	expectedNamespaceName := _ExceptionAdsReporter.NamespaceName,
	expectedClassName := 'LongDateTimeAssertionContext',
	expectedSize := XSIZEOF(_MetadataLongDateTimeAssertionContext),
	expectedAddress := ADR(_MetadataLongDateTimeAssertionContext)
);
assertObjectMetadata(
	object := _MetadataLongRealAssertionContext,
	expectedNamespaceName := _ExceptionAdsReporter.NamespaceName,
	expectedClassName := 'LongRealAssertionContext',
	expectedSize := XSIZEOF(_MetadataLongRealAssertionContext),
	expectedAddress := ADR(_MetadataLongRealAssertionContext)
);
assertObjectMetadata(
	object := _MetadataLongTimeAssertionContext,
	expectedNamespaceName := _ExceptionAdsReporter.NamespaceName,
	expectedClassName := 'LongTimeAssertionContext',
	expectedSize := XSIZEOF(_MetadataLongTimeAssertionContext),
	expectedAddress := ADR(_MetadataLongTimeAssertionContext)
);
assertObjectMetadata(
	object := _MetadataLongTimeOfDayAssertionContext,
	expectedNamespaceName := _ExceptionAdsReporter.NamespaceName,
	expectedClassName := 'LongTimeOfDayAssertionContext',
	expectedSize := XSIZEOF(_MetadataLongTimeOfDayAssertionContext),
	expectedAddress := ADR(_MetadataLongTimeOfDayAssertionContext)
);
assertObjectMetadata(
	object := _MetadataLWordAssertionContext,
	expectedNamespaceName := _ExceptionAdsReporter.NamespaceName,
	expectedClassName := 'LWordAssertionContext',
	expectedSize := XSIZEOF(_MetadataLWordAssertionContext),
	expectedAddress := ADR(_MetadataLWordAssertionContext)
);
assertObjectMetadata(
	object := _MetadataPointerAssertionContext,
	expectedNamespaceName := _ExceptionAdsReporter.NamespaceName,
	expectedClassName := 'PointerAssertionContext',
	expectedSize := XSIZEOF(_MetadataPointerAssertionContext),
	expectedAddress := ADR(_MetadataPointerAssertionContext)
);
assertObjectMetadata(
	object := _MetadataRealAssertionContext,
	expectedNamespaceName := _ExceptionAdsReporter.NamespaceName,
	expectedClassName := 'RealAssertionContext',
	expectedSize := XSIZEOF(_MetadataRealAssertionContext),
	expectedAddress := ADR(_MetadataRealAssertionContext)
);
assertObjectMetadata(
	object := _MetadataSIntAssertionContext,
	expectedNamespaceName := _ExceptionAdsReporter.NamespaceName,
	expectedClassName := 'SIntAssertionContext',
	expectedSize := XSIZEOF(_MetadataSIntAssertionContext),
	expectedAddress := ADR(_MetadataSIntAssertionContext)
);
assertObjectMetadata(
	object := _MetadataStringAssertionContext,
	expectedNamespaceName := _ExceptionAdsReporter.NamespaceName,
	expectedClassName := 'StringAssertionContext',
	expectedSize := XSIZEOF(_MetadataStringAssertionContext),
	expectedAddress := ADR(_MetadataStringAssertionContext)
);
assertObjectMetadata(
	object := _MetadataTimeAssertionContext,
	expectedNamespaceName := _ExceptionAdsReporter.NamespaceName,
	expectedClassName := 'TimeAssertionContext',
	expectedSize := XSIZEOF(_MetadataTimeAssertionContext),
	expectedAddress := ADR(_MetadataTimeAssertionContext)
);
assertObjectMetadata(
	object := _MetadataTimeOfDayAssertionContext,
	expectedNamespaceName := _ExceptionAdsReporter.NamespaceName,
	expectedClassName := 'TimeOfDayAssertionContext',
	expectedSize := XSIZEOF(_MetadataTimeOfDayAssertionContext),
	expectedAddress := ADR(_MetadataTimeOfDayAssertionContext)
);
assertObjectMetadata(
	object := _MetadataUDIntAssertionContext,
	expectedNamespaceName := _ExceptionAdsReporter.NamespaceName,
	expectedClassName := 'UDIntAssertionContext',
	expectedSize := XSIZEOF(_MetadataUDIntAssertionContext),
	expectedAddress := ADR(_MetadataUDIntAssertionContext)
);
assertObjectMetadata(
	object := _MetadataUIntAssertionContext,
	expectedNamespaceName := _ExceptionAdsReporter.NamespaceName,
	expectedClassName := 'UIntAssertionContext',
	expectedSize := XSIZEOF(_MetadataUIntAssertionContext),
	expectedAddress := ADR(_MetadataUIntAssertionContext)
);
assertObjectMetadata(
	object := _MetadataULIntAssertionContext,
	expectedNamespaceName := _ExceptionAdsReporter.NamespaceName,
	expectedClassName := 'ULIntAssertionContext',
	expectedSize := XSIZEOF(_MetadataULIntAssertionContext),
	expectedAddress := ADR(_MetadataULIntAssertionContext)
);
assertObjectMetadata(
	object := _MetadataUSIntAssertionContext,
	expectedNamespaceName := _ExceptionAdsReporter.NamespaceName,
	expectedClassName := 'USIntAssertionContext',
	expectedSize := XSIZEOF(_MetadataUSIntAssertionContext),
	expectedAddress := ADR(_MetadataUSIntAssertionContext)
);
assertObjectMetadata(
	object := _MetadataWideStringAssertionContext,
	expectedNamespaceName := _ExceptionAdsReporter.NamespaceName,
	expectedClassName := 'WideStringAssertionContext',
	expectedSize := XSIZEOF(_MetadataWideStringAssertionContext),
	expectedAddress := ADR(_MetadataWideStringAssertionContext)
);
assertObjectMetadata(
	object := _MetadataWordAssertionContext,
	expectedNamespaceName := _ExceptionAdsReporter.NamespaceName,
	expectedClassName := 'WordAssertionContext',
	expectedSize := XSIZEOF(_MetadataWordAssertionContext),
	expectedAddress := ADR(_MetadataWordAssertionContext)
);

first := _MetadataBoolAssertionContext;
second := _OtherBoolContext;
expect(condition := first.Equals(other := first), message := 'A context equals itself');
expectFalse(condition := first.Equals(other := second), message := 'Equal snapshots do not merge context identity');
expectFalse(condition := first.Equals(other := 0), message := 'A context is distinct from null');

group := _Runner.Empty;
expect(condition := group.ClassName <> '', message := 'A concrete group provides its class name');
expect(
	condition := group.NamespaceName = _Runner.NamespaceName,
	message := 'Group and runner share the consumer namespace'
);
expect(condition := group.SelfSize = XSIZEOF(_Runner.Empty), message := 'Group size includes its concrete storage');
expect(
	condition := group.SelfAddress = ADR(_Runner.Empty),
	message := 'Group identity points to the concrete instance'
);

named := _Runner.Empty;
displayName REF= named.Name;
concreteDisplayName REF= _Runner.Empty.Name;
expect(condition := __ISVALIDREF(displayName), message := 'INamed provides a valid name reference');
expect(condition := ADR(displayName) = ADR(concreteDisplayName), message := 'INamed borrows the same name storage');
expect(condition := displayName = "Empty", message := 'INamed exposes the constructor-copied group name');

checkContextObjects := TRUE;
END_METHOD

(*!
<summary>Checks deadline completion, BUSY failure termination and mutation guards.</summary>
<description>
Configures the persistent output leaf through a local reference without copying it.
The first run must exercise active mutation guards before the deadline. The second injects a BUSY failure.
Returns TRUE when all observations for this scenario are complete.
</description>
*)
METHOD PRIVATE checkDeadline : BOOL
VAR
	deadlineProbe : REFERENCE TO AssertionIsolationProbe;
	exceptionCode : __SYSTEM.ExceptionCode;
	rejected : BOOL;
	actualParent : TOF_Testing.ITestElement;
END_VAR
deadlineProbe REF= _DeadlineRun.DeadlineGroup.Child;

IF NOT _DeadlineConfigured THEN
	deadlineProbe.CompleteAfterCycle := 0;
	deadlineProbe.Timeout := T#1MS;
	_DeadlineRun.Reporter := _DeadlineReport;
	_DeadlineConfigured := TRUE;
END_IF

_DeadlineRun.Execute(cleanupTaskMemory := FALSE);
_DeadlineCalls := _DeadlineCalls + 1;

IF deadlineProbe.IsRunning AND_THEN NOT _DeadlineBusyFailureRun AND_THEN NOT _ActiveConfigurationChecked THEN

	__TRY
		deadlineProbe.Timeout := T#2S;
	__CATCH(exceptionCode)
		assertCaughtExceptionType(
			exceptionCode := exceptionCode,
			expectedTypeName := 'StandardException'
		);
		rejected := TRUE;
	__ENDTRY

	expect(condition := rejected, message := 'An active deadline cannot be changed');
	expect(
		condition := deadlineProbe.Timeout = T#1MS,
		message := 'Rejected mutation preserves the deadline'
	);
	_DeadlineRun.Reset();
	expect(
		condition := deadlineProbe.IsRunning AND_THEN NOT _DeadlineRun.IsFinished,
		message := 'Active Reset leaves the pending leaf running'
	);
	rejected := FALSE;

	__TRY
		_DeadlineRun.Reporter := _DeadlineReport;
	__CATCH(exceptionCode)
		assertCaughtExceptionType(
			exceptionCode := exceptionCode,
			expectedTypeName := 'StandardException'
		);
		rejected := TRUE;
	__ENDTRY

	expect(condition := rejected, message := 'Active runner rejects Reporter mutation');
	actualParent := deadlineProbe.Parent;
	expect(
		condition := actualParent = _DeadlineRun.Children[0],
		message := 'The active leaf retains its constructor-assigned parent'
	);
	_ActiveConfigurationChecked := TRUE;
END_IF

IF NOT _DeadlineRun.IsFinished AND_THEN _DeadlineCalls < _DeadlineScanLimit THEN
	RETURN;
END_IF

IF NOT _DeadlineBusyFailureRun THEN
	expect(condition := _DeadlineRun.IsFinished, message := 'A one-millisecond nominal deadline terminates');
	expect(condition := _ActiveConfigurationChecked, message := 'Deadline run exercises the active mutation guards');
	expectDInt(expected := 1, actual := _DeadlineRun.FailedTests, message := 'Deadline is one failed leaf');
	expectUDInt(
		expected := 1,
		actual := deadlineProbe.TeardownCalls,
		message := 'Deadline cleanup occurs once'
	);

	IF _DeadlineRun.IsFinished THEN
		_DeadlineBusyFailureRun := TRUE;
		_DeadlineCalls := 0;
		_DeadlineRun.Reset();
		deadlineProbe.Timeout := T#0S;
		deadlineProbe.FailSelfWhileBusy := TRUE;
		RETURN;
	END_IF
ELSE
	expect(condition := _DeadlineRun.IsFinished, message := 'A failed BUSY step terminates immediately');
	expectDInt(expected := 1, actual := _DeadlineRun.FailedTests, message := 'BUSY failure counts once');
	expectUDInt(
		expected := 1,
		actual := deadlineProbe.BodyCalls,
		message := 'Failed BUSY step does not run another body cycle'
	);
	expectUDInt(
		expected := 1,
		actual := deadlineProbe.TeardownCalls,
		message := 'Failed BUSY cleanup occurs once'
	);
END_IF

checkDeadline := TRUE;
END_METHOD

(*!
<summary>Checks copied native, fallback and long diagnostics after earlier task-cycle cleanup.</summary>
<description>
Requires the inner run to finish and publish its report before the suite accepts the diagnostic results.
Returns TRUE when all observations for this scenario are complete.
</description>
*)
METHOD PRIVATE checkDiagnostics : BOOL
VAR
	probe : REFERENCE TO DiagnosticProbe;
END_VAR
IF NOT _DiagnosticConfigured THEN
	probe REF= _DiagnosticRun.NativeDiagnostic;
	probe.ThrowNative := TRUE;
	probe REF= _DiagnosticRun.FormatterDiagnostic;
	probe.ThrowOnGetMessage := TRUE;
	_DiagnosticRun.Reporter := _DiagnosticReport;
	_DiagnosticConfigured := TRUE;
END_IF

_DiagnosticRun.Execute(cleanupTaskMemory := FALSE);
_DiagnosticCalls := _DiagnosticCalls + 1;

IF NOT _DiagnosticRun.IsFinished AND_THEN _DiagnosticCalls < 16 THEN
	RETURN;
END_IF

expect(condition := _DiagnosticRun.IsFinished, message := 'The diagnostic run finishes within 16 scans');
expect(condition := _DiagnosticReport.IsReady, message := 'The diagnostic report is complete');
expectDInt(
	expected := 3,
	actual := _DiagnosticRun.FailedTests,
	message := 'All injected errors are failed leaves'
);
expect(
	condition := TOF_Core.WideStrings.Contains(stringToSearchIn := _DiagnosticRun.NativeDiagnostic.FailureMessage,
		stringToFind := "ExecuteTest"),
	message := 'Native diagnostic has the interrupted stage'
);
expect(
	condition := TOF_Core.WideStrings.Contains(stringToSearchIn := _DiagnosticRun.FormatterDiagnostic.FailureMessage,
		stringToFind := "diagnostic unavailable"),
	message := 'Failing GetMessage retains stage/code fallback'
);
expect(
	condition := TOF_Core.WideStrings.Contains(stringToSearchIn := _DiagnosticRun.LongDiagnostic.FailureMessage,
		stringToFind := "END_OF_LONG_DIAGNOSTIC"),
	message := 'Long copied exception message is not narrowed to 255'
);
expectUDInt(
	expected := 1,
	actual := _DiagnosticRun.FormatterDiagnostic.TeardownCalls,
	message := 'Fallback still tears down once'
);
checkDiagnostics := TRUE;
END_METHOD

(*!
<summary>Checks a zero-child runner completes successfully with zero tests.</summary>
<description>Returns TRUE when all observations for this scenario are complete.</description>
*)
METHOD PRIVATE checkEmptyRun : BOOL
IF NOT _EmptyConfigured THEN
	_EmptyRun.Reporter := _EmptyReport;
	_EmptyConfigured := TRUE;
END_IF

_EmptyRun.Execute(cleanupTaskMemory := FALSE);
_EmptyCalls := _EmptyCalls + 1;

IF NOT _EmptyRun.IsFinished AND_THEN _EmptyCalls < _EmptyScanLimit THEN
	RETURN;
END_IF

expect(condition := _EmptyRun.IsFinished, message := 'An empty run must finish within the scan limit');
expect(condition := _EmptyRun.AllPassed, message := 'An empty run passes');
expectDInt(expected := 0, actual := _EmptyRun.TotalTests, message := 'No synthetic empty test');
checkEmptyRun := TRUE;
END_METHOD

(*!
<summary>Checks missing static storage, safe abort recovery rejection and invalid reporter outcomes.</summary>
<description>Returns TRUE when all observations for this scenario are complete.</description>
*)
METHOD PRIVATE checkExceptionClasses : BOOL
VAR
	exceptionCode : __SYSTEM.ExceptionCode;
	rejected : BOOL;
	diagnostic : TOF_Core.ERROR_MESSAGE;
END_VAR
__TRY
	_MissingConfigurationGroup.Reset(reporter := 0);
__CATCH(exceptionCode)
	assertCaughtExceptionType(exceptionCode := exceptionCode, expectedTypeName := 'DataMemberNotSpecifiedException');
	rejected := TRUE;
__ENDTRY

expect(condition := rejected, message := 'Group Reset rejects missing child-array storage');
_MissingConfigurationRunner.Execute(cleanupTaskMemory := FALSE);
expectDInt(
	expected := -1,
	actual := _MissingConfigurationRunner.ExitCode,
	message := 'Missing runner storage aborts'
);
assertCaughtExceptionType(
	exceptionCode := _MissingConfigurationRunner.CallbackException,
	expectedTypeName := 'DataMemberNotSpecifiedException'
);
rejected := FALSE;

__TRY
	_MissingConfigurationRunner.Reset();
__CATCH(exceptionCode)
	assertCaughtExceptionType(exceptionCode := exceptionCode, expectedTypeName := 'DataMemberNotSpecifiedException');
	rejected := TRUE;
__ENDTRY

expect(condition := rejected, message := 'Recovery rejects missing storage before any child access');
expectDInt(
	expected := -1,
	actual := _MissingConfigurationRunner.ExitCode,
	message := 'Invalid recovery retains abort'
);
rejected := FALSE;

__TRY
	_ExceptionAdsReporter.ReportTestCaseResult(
		groupPath := "",
		testName := "Invalid ADS outcome",
		outcome := TOF_Testing.TEST_OUTCOME.RUNNING,
		duration := T#0S,
		message := diagnostic
	);
__CATCH(exceptionCode)
	assertCaughtExceptionType(exceptionCode := exceptionCode, expectedTypeName := 'ArgumentValueNotSupportedException');
	rejected := TRUE;
__ENDTRY

expect(condition := rejected, message := 'Reporter rejects the actual nonterminal enum value');
checkExceptionClasses := TRUE;
END_METHOD

(*!
<summary>Verifies first-failure summary retention and per-run reset through the ADS reporter callbacks.</summary>
<description>Checks rejected writes, bounded ADS output for a root leaf, and reset on the next run.
Returns TRUE when all observations for this scenario are complete.
</description>
*)
METHOD PRIVATE checkAdsReporterSummary : BOOL
VAR
	diagnostic : TOF_Core.ERROR_MESSAGE;
END_VAR
_AdsSummaryReporter.ReportRunStart(testCount := 2);
_AdsSummaryReporter.RejectWrites := TRUE;
diagnostic := "Synthetic first diagnostic";
_AdsSummaryReporter.ReportTestCaseResult(
	groupPath := "Reporter regression",
	testName := "First leaf",
	outcome := TOF_Testing.TEST_OUTCOME.FAILED,
	duration := T#0S,
	message := diagnostic
);

_AdsSummaryReporter.RejectWrites := FALSE;
diagnostic := "Synthetic second diagnostic";
_AdsSummaryReporter.ReportTestCaseResult(
	groupPath := "Reporter regression",
	testName := "Second leaf",
	outcome := TOF_Testing.TEST_OUTCOME.FAILED,
	duration := T#0S,
	message := diagnostic
);

_AdsSummaryReporter.ReportRunEnd(
	totalTests := 2,
	passedTests := 0,
	failedTests := 2,
	skippedTests := 0,
	duration := T#0S
);

expect(
	condition := _AdsSummaryReporter.LastRunSummary =
		"[TOF_Testing] Finished: 0 passed, 2 failed, 0 skipped | First failure: First leaf: Synthetic first diagnostic",
	message := 'A second failure must preserve the first failure in the summary'
);

expect(
	condition := _AdsSummaryReporter.AcceptedMessage =
		"[TOF_Testing] Finished: 0 passed, 2 failed, 0 skipped | First failed test: First leaf",
	message := 'The completion record must identify the first failure even after its detail write is rejected'
);
expect(
	condition := _AdsSummaryReporter.FailedLogWriteCount = 1,
	message := 'Exactly one rejected write must be counted'
);
expect(
	condition := _AdsSummaryReporter.LastLogFailureMessage =
		"[TOF_Testing] Reporter regression/First leaf: Synthetic first diagnostic",
	message := 'Later accepted writes must preserve the rejected message'
);

_AdsSummaryReporter.ReportRunStart(testCount := 0);

expect(
	condition := _AdsSummaryReporter.LastRunSummary = "",
	message := 'Starting a new run must clear the retained summary'
);
expect(
	condition := _AdsSummaryReporter.FailedLogWriteCount = 0 AND_THEN _AdsSummaryReporter.LastLogFailureMessage = "",
	message := 'A successful start must clear earlier failed-write observations'
);

_AdsSummaryReporter.ReportRunEnd(
	totalTests := 0,
	passedTests := 0,
	failedTests := 0,
	skippedTests := 0,
	duration := T#0S
);

expect(
	condition := _AdsSummaryReporter.LastRunSummary = "[TOF_Testing] Finished: 0 passed, 0 failed, 0 skipped",
	message := 'An empty run must omit the earlier failure'
);

_AdsSummaryReporter.ReportRunStart(testCount := 1);
diagnostic := "Long diagnostic containing a literal %s. ";
TOF_Core.WideStrings.AppendFit255(
	diagnostic,
	"AAAAAAAAAAAAAAAAAAAAAAAAAAAAAAAAAAAAAAAAAAAAAAAAAAAAAAAAAAAAAAAAAAAAAAAAAAAAAAAA",
	"BBBBBBBBBBBBBBBBBBBBBBBBBBBBBBBBBBBBBBBBBBBBBBBBBBBBBBBBBBBBBBBBBBBBBBBBBBBBBBBB",
	"CCCCCCCCCCCCCCCCCCCCCCCCCCCCCCCCCCCCCCCCCCCCCCCCCCCCCCCCCCCCCCCCCCCCCCCCCCCCCCCC"
);
_AdsSummaryReporter.ReportTestCaseResult(
	groupPath := "",
	testName := "Long failure",
	outcome := TOF_Testing.TEST_OUTCOME.FAILED,
	duration := T#0S,
	message := diagnostic
);

expect(
	condition := TOF_Core.WideStrings.GetLength(value := _AdsSummaryReporter.AcceptedMessage) = 200,
	message := 'A long ADS diagnostic must fit within the reporter limit'
);
expect(
	condition := Tc2_Standard.WLEFT(STR := _AdsSummaryReporter.AcceptedMessage, SIZE := 27) =
		"[TOF_Testing] Long failure:",
	message := 'A root leaf is logged without a leading group separator'
);

_AdsSummaryReporter.RejectWrites := TRUE;
_AdsSummaryReporter.ReportRunEnd(
	totalTests := 1,
	passedTests := 0,
	failedTests := 1,
	skippedTests := 0,
	duration := T#0S
);
expect(
	condition := _AdsSummaryReporter.LastLogFailureMessage =
		"[TOF_Testing] Finished: 0 passed, 1 failed, 0 skipped | First failed test: Long failure",
	message := 'Rejection must retain the exact completion record independently of diagnostic length'
);
expect(
	condition := _AdsSummaryReporter.FailedLogWriteCount = 1,
	message := 'A rejected completion record must be counted once'
);
_AdsSummaryReporter.RejectWrites := FALSE;

checkAdsReporterSummary := TRUE;
END_METHOD

(*!
<summary>Recovers a throwing external child, including a failed first recovery attempt.</summary>
<description>Explicitly releases the modeled resource before requesting reset recovery.
Returns TRUE when all observations for this scenario are complete.
</description>
*)
METHOD PRIVATE checkExternalRecovery : BOOL
VAR
	exceptionCode : __SYSTEM.ExceptionCode;
	rejected : BOOL;
	externalCase : REFERENCE TO ExternalElementProbe;
	actualParent : TOF_Testing.ITestElement;
END_VAR
IF NOT _ExternalConfigured THEN
	_ExternalRun.Reporter := _ExternalReport;
	_ExternalConfigured := TRUE;
END_IF

_ExternalRun.Execute(cleanupTaskMemory := FALSE);
_ExternalCalls := _ExternalCalls + 1;

IF NOT _ExternalRun.IsFinished THEN
	IF _ExternalCalls < 16 THEN
		RETURN;
	END_IF

	expect(condition := FALSE, message := 'The external recovery run must finish within 16 scans');
	_ExternalRun.ExternalCase.ReleaseResource();
	checkExternalRecovery := TRUE;

	RETURN;
END_IF

IF NOT _ExternalRecovered THEN
	expectDInt(expected := -1, actual := _ExternalRun.ExitCode, message := 'External child aborts');
	expect(
		condition := _ExternalRun.ExternalCase.ResourceActive,
		message := 'Abort does not silently release user resources'
	);
	_ExternalRun.Execute(cleanupTaskMemory := FALSE);
	expectUDInt(
		expected := 1,
		actual := _ExternalRun.ExternalCase.ExecuteCalls,
		message := 'The aborted callback is not retried before explicit recovery'
	);
	externalCase REF= _ExternalRun.ExternalCase;
	externalCase.ReleaseResource();
	expectFalse(
		condition := externalCase.ResourceActive,
		message := 'Explicit resource release completes before reset recovery'
	);
	externalCase.ThrowOnReset := TRUE;

	__TRY
		_ExternalRun.Reset();
	__CATCH(exceptionCode)
		assertCaughtExceptionType(
			exceptionCode := exceptionCode,
			expectedTypeName := 'StandardException'
		);
		rejected := TRUE;
	__ENDTRY

	expect(condition := rejected, message := 'Custom recovery Reset failure propagates');
	expectDInt(expected := -1, actual := _ExternalRun.ExitCode, message := 'Failed recovery retains abort');
	externalCase.ThrowOnReset := FALSE;
	externalCase.ThrowOnExecute := FALSE;
	_ExternalRun.Reset();
	actualParent := _ExternalRun.ExternalCase.Parent;
	expect(condition := actualParent = 0, message := 'The recovered root remains parentless');
	expectUDInt(
		expected := 3,
		actual := _ExternalRun.ExternalCase.ResetCalls,
		message := 'Failed reset was retried'
	);
	_ExternalRecovered := TRUE;
	_ExternalCalls := 0;
	RETURN;
END_IF

expect(condition := _ExternalRun.AllPassed, message := 'The same static tree succeeds after explicit recovery');
expectDInt(expected := 1, actual := _ExternalRun.PassedTests, message := 'The recovered root contributes one leaf');
expect(condition := _ExternalReport.IsReady, message := 'The recovered run completes its report');
expectUDInt(
	expected := 2,
	actual := _ExternalRun.ExternalCase.ExecuteCalls,
	message := 'Execute resumes only in the new run'
);
checkExternalRecovery := TRUE;
END_METHOD

(*!
<summary>Checks direct-child interface dispatch, fixed ordering and explicit accessor failures.</summary>
<description>
Borrows persistent fixtures before execution and after a rejected Reset. Test-only slot corruption is restored
before returning. Child identity is compared through ITestElement on both sides; indexed observation
invokes no child body.

Returns TRUE when all observations for this scenario are complete.
</description>
*)
METHOD PRIVATE checkIndexedChildren : BOOL
VAR
	element : TOF_Testing.ITestElement;
	parentElement : TOF_Testing.IParentTestElement;
	child : TOF_Testing.ITestElement;
	expectedChild : TOF_Testing.ITestElement;
	supportsChildren : BOOL;
	exceptionCode : __SYSTEM.ExceptionCode;
	rejected : BOOL;
	firstBodyCalls : UDINT;
END_VAR
element := _IndexedGroup;
supportsChildren := __QUERYINTERFACE(element, parentElement);
expect(condition := supportsChildren, message := 'A group exposes the direct-child capability');

IF NOT supportsChildren THEN
	checkIndexedChildren := TRUE;
	RETURN;
END_IF

firstBodyCalls := _IndexedGroup.First.BodyCalls;
expect(condition := parentElement.ChildCount = 2, message := 'The capability reports the fixed direct count');
expectedChild := _IndexedGroup.First;
child := parentElement.GetChildByIndex(index := 0);
expect(condition := child = expectedChild, message := 'Index zero borrows the first child');
expectedChild := _IndexedGroup.Second;
child := parentElement.GetChildByIndex(index := 1);
expect(condition := child = expectedChild, message := 'The last valid index borrows the last child');

__TRY
	child := parentElement.GetChildByIndex(index := 2);
__CATCH(exceptionCode)
	assertCaughtExceptionType(exceptionCode := exceptionCode, expectedTypeName := 'ArgumentOutOfRangeException');
	rejected := TRUE;
__ENDTRY

expect(condition := rejected, message := 'Index equal to ChildCount is rejected');
rejected := FALSE;

__TRY
	child := parentElement.GetChildByIndex(index := TOF_Core.SignedInt16.MAX_VALUE);
__CATCH(exceptionCode)
	assertCaughtExceptionType(exceptionCode := exceptionCode, expectedTypeName := 'ArgumentOutOfRangeException');
	rejected := TRUE;
__ENDTRY

expect(condition := rejected, message := 'The largest representable index is rejected before indexing');
parentElement := _Runner.Empty;
expect(condition := parentElement.ChildCount = TOF_Core.SignedInt16.ZERO, message := 'An empty group reports zero direct children');
rejected := FALSE;

__TRY
	child := parentElement.GetChildByIndex(index := 0);
__CATCH(exceptionCode)
	assertCaughtExceptionType(exceptionCode := exceptionCode, expectedTypeName := 'ArgumentOutOfRangeException');
	rejected := TRUE;
__ENDTRY

expect(condition := rejected, message := 'A valid empty array has no valid child index');
parentElement := _MissingConfigurationGroup;
rejected := FALSE;

__TRY
	child := parentElement.GetChildByIndex(index := TOF_Core.SignedInt16.MAX_VALUE);
__CATCH(exceptionCode)
	assertCaughtExceptionType(exceptionCode := exceptionCode, expectedTypeName := 'DataMemberNotSpecifiedException');
	rejected := TRUE;
__ENDTRY

expect(condition := rejected, message := 'Missing storage is diagnosed before an invalid index');

// A failed Reset does not prevent observing an existing slot; the missing selected slot remains an error.
_IndexedGroup.Children[1] := 0;
rejected := FALSE;

__TRY
	_IndexedGroup.Reset(reporter := 0);
__CATCH(exceptionCode)
	assertCaughtExceptionType(exceptionCode := exceptionCode, expectedTypeName := 'DataMemberNotSpecifiedException');
	rejected := TRUE;
__ENDTRY

expect(condition := rejected, message := 'The injected missing slot rejects Reset');
parentElement := _IndexedGroup;
expectedChild := _IndexedGroup.First;
child := parentElement.GetChildByIndex(index := 0);
expect(condition := child = expectedChild, message := 'An existing slot can be observed after failed Reset');
rejected := FALSE;

__TRY
	child := parentElement.GetChildByIndex(index := 1);
__CATCH(exceptionCode)
	assertCaughtExceptionType(exceptionCode := exceptionCode, expectedTypeName := 'DataMemberNotSpecifiedException');
	rejected := TRUE;
__ENDTRY

expect(condition := rejected, message := 'A null selected slot is a missing member');
_IndexedGroup.Children[1] := _IndexedGroup.Second;
expectUDInt(
	expected := firstBodyCalls,
	actual := _IndexedGroup.First.BodyCalls,
	message := 'Indexed observation invokes no child body'
);
_IndexedGroup.Reset(reporter := 0);
checkIndexedChildren := TRUE;
END_METHOD

(*!
<summary>Checks live root-to-element paths independently of Reset and reporting.</summary>
<description>
Checks interface dispatch, own-name inclusion, empty names, Unicode, root-prefix truncation and cycles among ancestors.
Synthetic parent-only chains isolate GetPath; they are never registered or executed as group compositions.
The existing nested and repeated-run cases independently check JUnit group paths without the leaf name.

Returns TRUE when all observations for this scenario are complete.
</description>
*)
METHOD PRIVATE checkPaths : BOOL
VAR
	element : TOF_Testing.ITestElement;
	named : TOF_Core.INamed;
	actualPath : WSTRING(255);
	expectedPath : WSTRING(255);
	exceptionCode : __SYSTEM.ExceptionCode;
	rejected : BOOL;
	diagnostic : TOF_Core.ERROR_MESSAGE;
	content : POINTER TO STRING;
	longName : WSTRING(81);
	expectedXmlName : STRING(255);
END_VAR
expectedPath := "AAAAAAAAAAAAAAAAAAAAAAAAAAAAAAAAAAAAAAAAAAAAAAAAAAAAAAAAAAAAAAAAAAAAAAAAAAAAAAAA";
named := _PathLongName;
expect(condition := named.Name = expectedPath, message := 'INamed retains the first 80 name characters');
actualPath := _PathLongName.GetPath();
expect(condition := actualPath = expectedPath, message := 'A root path observes the same bounded name');
longName := "AAAAAAAAAAAAAAAAAAAAAAAAAAAAAAAAAAAAAAAAAAAAAAAAAAAAAAAAAAAAAAAAAAAAAAAAAAAAAAAAB";
_PathReport.ReportRunStart(testCount := 1);
_PathReport.ReportTestCaseResult(
	groupPath := "",
	testName := longName,
	outcome := TOF_Testing.TEST_OUTCOME.PASSED,
	duration := T#0S,
	message := diagnostic
);
_PathReport.ReportRunEnd(totalTests := 1, passedTests := 1, failedTests := 0, skippedTests := 0, duration := T#0S);
content := _PathReport.ContentAddress;
expectedXmlName := TOF_Core.Strings.Concat255('name="', TO_STRING(expectedPath), '"');
expect(condition := _PathReport.IsReady AND_THEN content <> 0, message := 'The bounded-name report completes');

IF content <> 0 THEN
	expect(
		condition := TOF_Core.Strings.Contains(stringToSearchIn := content^, stringToFind := expectedXmlName),
		message := 'Reporter input retains exactly the first 80 name characters'
	);
END_IF

element := _DuplicateGroup;
actualPath := element.GetPath();
expect(condition := actualPath = "Duplicates", message := 'A root path contains its own name');
actualPath := _DuplicateGroup.First.GetPath();
expect(condition := actualPath = "Duplicates/First", message := 'A child path includes its group and own name');
actualPath := _Runner.FailureOuter.Failures.BodyFailure.GetPath();
expect(
	condition := actualPath = "Nested/Failures/Body failure",
	message := 'Ancestor names are ordered from the root'
);
actualPath := _Runner.Pass.GetPath();
expect(condition := actualPath = "", message := 'A nameless root has an empty path');
actualPath := _PathEmpty.GetPath();
expectedPath := "AAAAAAAAAAAAAAAAAAAAAAAAAAAAAAAAAAAAAAAAAAAAAAAAAAAAAAAAAAAAAAAAAAAAAAAAAAAAAAAA";
expect(condition := actualPath = expectedPath, message := 'An empty own name adds no separator');
actualPath := _PathUnicode.GetPath();
expectedPath := "AAAAAAAAAAAAAAAAAAAAAAAAAAAAAAAAAAAAAAAAAAAAAAAAAAAAAAAAAAAAAAAAAAAAAAAAAAAAAAAA/Ω";
expect(condition := actualPath = expectedPath, message := 'Empty ancestors are skipped and Unicode is preserved');
actualPath := _PathFourth.GetPath();
expectedPath := Tc2_Utilities.WCONCAT(
	STR1 := "AAAAAAAAAAAAAAAAAAAAAAAAAAAAAAAAAAAAAAAAAAAAAAAAAAAAAAAAAAAAAAAAAAAAAAAAAAAAAAAA/",
	STR2 := "BBBBBBBBBBBBBBBBBBBBBBBBBBBBBBBBBBBBBBBBBBBBBBBBBBBBBBBBBBBBBBBBBBBBBBBBBBBBBBBB/"
);
expectedPath := Tc2_Utilities.WCONCAT(
	STR1 := expectedPath,
	STR2 := "CCCCCCCCCCCCCCCCCCCCCCCCCCCCCCCCCCCCCCCCCCCCCCCCCCCCCCCCCCCCCCCCCCCCCCCCCCCCCCCC/DDDDDDDDDDD…"
);
expect(condition := actualPath = expectedPath, message := 'Overflow retains the root prefix and final ellipsis');

__TRY
	actualPath := _ParentGroup.Child.GetPath();
__CATCH(exceptionCode)
	assertCaughtExceptionType(exceptionCode := exceptionCode, expectedTypeName := 'StandardException');
	rejected := TRUE;
__ENDTRY

expect(condition := rejected, message := 'A cycle among ancestors is rejected without endless traversal');
actualPath := _ReportPathInner.GetPath();
_PathReport.ReportRunStart(testCount := 1);
_PathReport.ReportTestCaseResult(
	groupPath := actualPath,
	testName := "Leaf",
	outcome := TOF_Testing.TEST_OUTCOME.PASSED,
	duration := T#0S,
	message := diagnostic
);
_PathReport.ReportRunEnd(totalTests := 1, passedTests := 1, failedTests := 0, skippedTests := 0, duration := T#0S);
content := _PathReport.ContentAddress;
expect(condition := _PathReport.IsReady AND_THEN content <> 0, message := 'The deep-path report completes');

IF content <> 0 THEN
	expect(
		condition := TOF_Core.Strings.Contains(
			stringToSearchIn := content^,
			stringToFind := 'name="Leaf" classname="Report root/Middle/Inner"'
		),
		message := 'JUnit preserves all three group ancestors and keeps the leaf name separate'
	);
END_IF

checkPaths := TRUE;
END_METHOD

(*!
<summary>Verifies that a reporter failure aborts once after teardown and clears the reporter reference.</summary>
<description>The same leaf runs with a replacement reporter after a completed abort and Reset.
An incomplete run fails when it reaches the scan limit. Returns TRUE when the scenario has an outcome.
</description>
*)
METHOD PRIVATE checkReporterAbort : BOOL
VAR
	exceptionCode : __SYSTEM.ExceptionCode;
	rejected : BOOL;
	diagnostic : TOF_Core.ERROR_MESSAGE;
	actualParent : TOF_Testing.ITestElement;
END_VAR
IF _AbortRecovered THEN
	_AbortRun.Execute(cleanupTaskMemory := FALSE);
	_AbortCalls := _AbortCalls + 1;

	IF NOT _AbortRun.IsFinished AND_THEN _AbortCalls < 16 THEN
		RETURN;
	END_IF

	expect(condition := _AbortRun.IsFinished, message := 'The recovered reporter run finishes within 16 scans');
	expect(condition := _AbortRun.IsFinished AND_THEN _AbortRun.AllPassed,
		message := 'The same static tree passes after reporter abort');
	expectUDInt(
		expected := 1,
		actual := _AbortRun.AbortCase.BodyCalls,
		message := 'The same root executes once in the new run'
	);
	expectUDInt(expected := 1, actual := _AbortReport.ResultCalls, message := 'Old reporter is not retried');
	checkReporterAbort := TRUE;
	RETURN;
END_IF

IF NOT _AbortConfigured THEN

	__TRY
		_InvalidReport.ReportTestCaseResult(
			groupPath := "",
			testName := "Invalid outcome",
			outcome := TOF_Testing.TEST_OUTCOME.NOT_RUN,
			duration := T#0S,
			message := diagnostic
		);
	__CATCH(exceptionCode)
		assertCaughtExceptionType(
			exceptionCode := exceptionCode,
			expectedTypeName := 'ArgumentValueNotSupportedException'
		);
		rejected := TRUE;
	__ENDTRY

	expect(condition := rejected, message := 'A reporter rejects a nonterminal outcome');
	_AbortRun.Reporter := _AbortReport;
	_AbortConfigured := TRUE;
END_IF

_AbortRun.Execute(cleanupTaskMemory := FALSE);
_AbortCalls := _AbortCalls + 1;

IF NOT _AbortRun.IsFinished THEN
	IF _AbortCalls < 16 THEN
		RETURN;
	END_IF

	expect(condition := FALSE, message := 'Callback abort must terminate within 16 scans');
	checkReporterAbort := TRUE;

	RETURN;
END_IF

IF _AbortPostCalls < 2 THEN
	_AbortPostCalls := _AbortPostCalls + 1;
	RETURN;
END_IF

expectDInt(expected := -1, actual := _AbortRun.ExitCode, message := 'Callback abort has a distinct exit code');
expectUDInt(expected := 1, actual := _AbortReport.ResultCalls, message := 'The callback is never retried');
expectUDInt(
	expected := 1,
	actual := _AbortRun.AbortCase.TeardownCalls,
	message := 'Cleanup precedes result reporting'
);
expect(
	condition := _AbortRun.AbortCase.IsFinished AND_THEN _AbortRun.AbortCase.Reporter = 0,
	message := 'A completed leaf clears its reporter reference even when result delivery throws'
);
expectFalse(condition := _AbortReport.IsReady, message := 'An aborted report remains incomplete');
expect(
	condition := TOF_Core.WideStrings.Contains(stringToSearchIn := _AbortRun.CallbackMessage,
		stringToFind := "Reporter failed"),
	message := 'External callback diagnostic is copied'
);
_AbortRun.Reset();
expect(condition := _AbortRun.CallbackMessage = "", message := 'Reset clears copied callback diagnostic');
actualParent := _AbortRun.AbortCase.Parent;
expect(condition := actualParent = 0, message := 'The same root remains parentless after recovery');
_AbortRun.Reporter := _AbortRecoveryReport;
_AbortRecovered := TRUE;
_AbortCalls := 0;
END_METHOD

(*!
<summary>Checks static root validation, recovery guards and absence of cyclic topology scans.</summary>
<description>Deliberately corrupts test-only slots, restoring them before valid recovery and before execution reaches them.
Returns TRUE when all observations for this scenario are complete.
</description>
*)
METHOD PRIVATE checkRunnerTopology : BOOL
VAR
	exceptionCode : __SYSTEM.ExceptionCode;
	rejected : BOOL;
	runningRoot : REFERENCE TO AssertionIsolationProbe;
	actualParent : TOF_Testing.ITestElement;
END_VAR
IF NOT _RootTopologyConfigured THEN
	_RootTopologyRunner.Reporter := _RootTopologyReport;
	_RootTopologyRunner.RootTopologyFirst.Reset(reporter := 0);
	_RootTopologyRunner.RootTopologyFirst.Execute();
	_RootTopologyRunner.Children[1] := 0;
	_RootTopologyRunner.Execute(cleanupTaskMemory := FALSE);
	expectDInt(expected := -1, actual := _RootTopologyRunner.ExitCode, message := 'A null root aborts startup');
	assertCaughtExceptionType(
		exceptionCode := _RootTopologyRunner.CallbackException,
		expectedTypeName := 'DataMemberNotSpecifiedException'
	);
	expect(
		condition := _RootTopologyRunner.RootTopologyFirst.IsFinished,
		message := 'All direct roots are validated before the first Reset'
	);
	expectFalse(condition := _RootTopologyReport.IsReady, message := 'Invalid startup produces no completed report');
	expect(
		condition := _RootTopologyReport.ContentLength = TOF_Core.UnsignedInt32.ZERO,
		message := 'Invalid startup does not call ReportRunStart'
	);
	rejected := FALSE;

	__TRY
		_RootTopologyRunner.Reset();
	__CATCH(exceptionCode)
		assertCaughtExceptionType(exceptionCode := exceptionCode, expectedTypeName := 'DataMemberNotSpecifiedException');
		rejected := TRUE;
	__ENDTRY

	expect(condition := rejected, message := 'Recovery validates slots before dereferencing an invalid tree');
	expectDInt(
		expected := -1,
		actual := _RootTopologyRunner.ExitCode,
		message := 'Failed recovery retains abort'
	);
	_RootTopologyRunner.Children[1] := _RootTopologyRunner.RootTopologyGroup;
	_RootTopologyRunner.Reset();
	_RootTopologyRunner.Children[1] := _RootTopologyRunner.RootTopologyFirst;
	_RootTopologyRunner.Execute(cleanupTaskMemory := FALSE);
	expectDInt(
		expected := -1,
		actual := _RootTopologyRunner.ExitCode,
		message := 'Duplicate roots abort startup'
	);
	assertCaughtExceptionType(exceptionCode := _RootTopologyRunner.CallbackException, expectedTypeName := 'StandardException');
	_RootTopologyRunner.Children[1] := _RootTopologyRunner.RootTopologyGroup;
	_RootTopologyRunner.Reset();
	_RootTopologyRunner.Children[0] := _RootTopologyRunner.RootTopologyGroup.Child;
	_RootTopologyRunner.Execute(cleanupTaskMemory := FALSE);
	expectDInt(
		expected := -1,
		actual := _RootTopologyRunner.ExitCode,
		message := 'A group-owned root aborts startup'
	);
	assertCaughtExceptionType(exceptionCode := _RootTopologyRunner.CallbackException, expectedTypeName := 'StandardException');
	_RootTopologyRunner.Children[0] := _RootTopologyRunner.RootTopologyFirst;
	_RootTopologyRunner.Reset();
	_RootTopologyRunner.RootTopologyFirst.Execute();
	_RootTopologyRunner.Children[1] := _Runner.FailureOuter.Failures;
	_RootTopologyRunner.Execute(cleanupTaskMemory := FALSE);
	expectDInt(
		expected := -1,
		actual := _RootTopologyRunner.ExitCode,
		message := 'A nested group cannot also occupy a root slot'
	);
	assertCaughtExceptionType(exceptionCode := _RootTopologyRunner.CallbackException, expectedTypeName := 'StandardException');
	expect(
		condition := _RootTopologyRunner.RootTopologyFirst.IsFinished,
		message := 'Owned-group rejection occurs before the first direct Reset'
	);
	expect(
		condition := _RootTopologyReport.ContentLength = TOF_Core.UnsignedInt32.ZERO,
		message := 'Owned-group rejection does not start reporting'
	);
	rejected := FALSE;

	__TRY
		_RootTopologyRunner.Reset();
	__CATCH(exceptionCode)
		assertCaughtExceptionType(exceptionCode := exceptionCode, expectedTypeName := 'StandardException');
		rejected := TRUE;
	__ENDTRY

	expect(condition := rejected, message := 'Abort recovery also rejects a group-owned root');
	expectDInt(expected := -1, actual := _RootTopologyRunner.ExitCode, message := 'Invalid recovery retains abort');
	_RootTopologyRunner.Children[1] := _RootTopologyRunner.RootTopologyGroup;
	_RootTopologyRunner.Reset();
	runningRoot REF= _RootTopologyRunner.RunningRoot;
	runningRoot.Timeout := T#0S;
	_RootTopologyRunner.RunningRoot.Reset(reporter := 0);
	_RootTopologyRunner.RunningRoot.Execute();
	expect(condition := _RootTopologyRunner.RunningRoot.IsRunning, message := 'The active-root fixture is pending');
	_RootTopologyRunner.Children[0] := _RootTopologyRunner.RunningRoot;
	_RootTopologyRunner.Execute(cleanupTaskMemory := FALSE);
	expectDInt(
		expected := -1,
		actual := _RootTopologyRunner.ExitCode,
		message := 'An active root aborts startup'
	);
	assertCaughtExceptionType(exceptionCode := _RootTopologyRunner.CallbackException, expectedTypeName := 'StandardException');
	_RootTopologyRunner.RunningRoot.Reset(reporter := 0);
	_RootTopologyRunner.Children[0] := _RootTopologyRunner.RootTopologyFirst;
	_RootTopologyRunner.Reset();
	_RootTopologyRunner.Execute(cleanupTaskMemory := FALSE);
	expectFalse(condition := _RootTopologyRunner.IsFinished, message := 'Valid startup prepares the static roots');

	// Fault injection: restore the unused slot immediately after driving the first root.
	_RootTopologyRunner.Children[1] := 0;
	_RootTopologyRunner.Execute(cleanupTaskMemory := FALSE);
	_RootTopologyRunner.Children[1] := _RootTopologyRunner.RootTopologyGroup;
	expectDInt(
		expected := 0,
		actual := _RootTopologyRunner.ExitCode,
		message := 'Execution does not rescan root slots'
	);
	_RootTopologyConfigured := TRUE;
END_IF

_RootTopologyRunner.Execute(cleanupTaskMemory := FALSE);
_RootTopologyCalls := _RootTopologyCalls + 1;

IF NOT _RootTopologyRunner.IsFinished AND_THEN _RootTopologyCalls < 16 THEN
	RETURN;
END_IF

expect(condition := _RootTopologyRunner.IsFinished, message := 'The topology run finishes within 16 scans');
expect(
	condition := _RootTopologyRunner.IsFinished AND_THEN _RootTopologyRunner.AllPassed,
	message := 'The owned static roots execute successfully'
);
expectDInt(
	expected := 2,
	actual := _RootTopologyRunner.PassedTests,
	message := 'Two direct or nested leaves pass'
);
expectUDInt(
	expected := 1,
	actual := _RootTopologyRunner.RootTopologyFirst.BodyCalls,
	message := 'The first root executes once in the valid run'
);
expectUDInt(
	expected := 1,
	actual := _RootTopologyRunner.RootTopologyGroup.Child.BodyCalls,
	message := 'The nested group executes its owned leaf'
);
actualParent := _RootTopologyRunner.RootTopologyFirst.Parent;
expect(condition := actualParent = 0, message := 'Runner roots remain parentless');
actualParent := _RootTopologyRunner.RootTopologyGroup.Child.Parent;
expect(
	condition := actualParent <> 0,
	message := 'A nested leaf retains its constructor-assigned parent'
);
checkRunnerTopology := TRUE;
END_METHOD

(*!
<summary>Checks fixed parents, missing or repeated children, parent mismatch, cycles, ordered dispatch and repeat execution.</summary>
<description>
Fault injection deliberately mutates a test-only array between rejected operations and briefly during execution
to detect redundant validation. Restore every unused slot before execution reaches it.

Returns TRUE when all observations for this scenario are complete.
</description>
*)
METHOD PRIVATE checkTopology : BOOL
VAR
	exceptionCode : __SYSTEM.ExceptionCode;
	rejected : BOOL;
	expectedParent : TOF_Testing.ITestElement;
	actualParent : TOF_Testing.ITestElement;
END_VAR
expectedParent := _DuplicateGroup;
actualParent := _DuplicateGroup.First.Parent;
expect(condition := actualParent = expectedParent, message := 'Parent is assigned at construction');
actualParent := _DuplicateGroup.Parent;
expect(condition := actualParent = 0, message := 'A root is constructed without a parent');

// Deliberately corrupt the borrowed test-only array to inject topology faults.
// A later execution probe restores its unused slot before that slot is reached.
_DuplicateGroup.Children[1] := 0;

__TRY
	_DuplicateGroup.Reset(reporter := 0);
__CATCH(exceptionCode)
	assertCaughtExceptionType(exceptionCode := exceptionCode, expectedTypeName := 'DataMemberNotSpecifiedException');
	rejected := TRUE;
__ENDTRY

expect(condition := rejected, message := 'A null fixed child is rejected by Reset');
expectUDInt(
	expected := 0,
	actual := _DuplicateGroup.First.BodyCalls,
	message := 'No earlier child body executes'
);
rejected := FALSE;
_DuplicateGroup.Children[1] := _DuplicateGroup.First;

__TRY
	_DuplicateGroup.Reset(reporter := 0);
__CATCH(exceptionCode)
	assertCaughtExceptionType(exceptionCode := exceptionCode, expectedTypeName := 'StandardException');
	rejected := TRUE;
__ENDTRY

expect(condition := rejected, message := 'Duplicate fixed slots are rejected');
rejected := FALSE;
_DuplicateGroup.Children[1] := _RootTopologyRunner.RootTopologyGroup.Child;

__TRY
	_DuplicateGroup.Reset(reporter := 0);
__CATCH(exceptionCode)
	assertCaughtExceptionType(exceptionCode := exceptionCode, expectedTypeName := 'StandardException');
	rejected := TRUE;
__ENDTRY

expect(condition := rejected, message := 'A child assigned to another group is rejected');
actualParent := _DuplicateGroup.First.Parent;
expect(condition := actualParent = expectedParent, message := 'Rejection never changes Parent');
_DuplicateGroup.Children[1] := _DuplicateGroup.Second;
rejected := FALSE;

__TRY
	_ParentGroup.Reset(reporter := 0);
__CATCH(exceptionCode)
	assertCaughtExceptionType(exceptionCode := exceptionCode, expectedTypeName := 'StandardException');
	rejected := TRUE;
__ENDTRY

expect(condition := rejected, message := 'A cycle assigned by constructors is rejected before recursion');

_DuplicateGroup.Reset(reporter := 0);
// Fault injection: an unused slot must not be rescanned in Execute; restore before that slot is reached.
_DuplicateGroup.Children[1] := 0;
_DuplicateGroup.Execute();
expectUDInt(
	expected := 1,
	actual := _DuplicateGroup.First.BodyCalls,
	message := 'The first Execute reaches the first owned child through Children'
);
expectUDInt(
	expected := 0,
	actual := _DuplicateGroup.Second.BodyCalls,
	message := 'The first Execute does not reach the second owned child'
);
_DuplicateGroup.Children[1] := _DuplicateGroup.Second;
_DuplicateGroup.Execute();
expect(condition := _DuplicateGroup.IsFinished, message := 'A valid static group finishes without Configure');
expectDInt(expected := 2, actual := _DuplicateGroup.PassedCount, message := 'Both owned leaves pass');
_DuplicateGroup.Reset(reporter := 0);
_DuplicateGroup.Execute();
_DuplicateGroup.Execute();
expectDInt(
	expected := 2,
	actual := _DuplicateGroup.PassedCount,
	message := 'Reset supports another fixed-tree run'
);
expectUDInt(
	expected := 1,
	actual := _DuplicateGroup.First.BodyCalls,
	message := 'A repeated leaf executes once'
);
actualParent := _DuplicateGroup.First.Parent;
expect(condition := actualParent = expectedParent, message := 'Repeated runs preserve Parent');
_DuplicateGroup.Children[1] := 0;
rejected := FALSE;

__TRY
	_DuplicateGroup.Reset(reporter := 0);
__CATCH(exceptionCode)
	assertCaughtExceptionType(exceptionCode := exceptionCode, expectedTypeName := 'DataMemberNotSpecifiedException');
	rejected := TRUE;
__ENDTRY

expect(condition := rejected, message := 'Invalid topology is rejected on a later Reset too');
expect(
	condition := _DuplicateGroup.First.IsFinished,
	message := 'Validation precedes the first direct child Reset'
);
_DuplicateGroup.Children[1] := _DuplicateGroup.Second;
checkTopology := TRUE;
END_METHOD

(*!
<summary>Checks long XML diagnostics, supplementary Unicode, isolated surrogates and XML controls.</summary>
<description>Returns TRUE when all observations for this scenario are complete.</description>
*)
METHOD PRIVATE checkXmlEncoding : BOOL
VAR
	diagnostic : TOF_Core.ERROR_MESSAGE;
	characters : POINTER TO WORD;
	content : POINTER TO STRING;
	i : UDINT;
END_VAR
// U+1F600 is a surrogate pair; it is followed by an isolated high surrogate, U+0001, TAB and ampersand.
characters := ADR(diagnostic);
characters[0] := 16#D83D;
characters[1] := 16#DE00;
characters[2] := 16#D800;
characters[3] := 16#0001;
characters[4] := 16#0009;
characters[5] := 16#0026;

FOR i := 6 TO 405 DO
	characters[i] := 16#0078;
END_FOR

characters[406] := TOF_Core.UnsignedInt16.MIN_VALUE;
TOF_Core.WideStrings.AppendFit(targetString := diagnostic, sourceString := "END_OF_XML_DIAGNOSTIC");
_XmlReport.ReportRunStart(testCount := 1);
_XmlReport.ReportTestCaseResult(
	groupPath := "Wide",
	testName := "",
	outcome := TOF_Testing.TEST_OUTCOME.FAILED,
	duration := T#1250MS,
	message := diagnostic
);
_XmlReport.ReportRunEnd(totalTests := 1, passedTests := 0, failedTests := 1, skippedTests := 0, duration := T#1250MS);
content := _XmlReport.ContentAddress;
expect(condition := _XmlReport.IsReady AND_THEN content <> 0, message := 'Completed Unicode XML has a buffer');

IF content <> 0 THEN
	expect(
		condition := TOF_Core.Strings.Contains(stringToSearchIn := content^,
			stringToFind := '&#128512;&#65533;&#65533;&#9;&amp;'),
		message := 'Surrogate pair, isolated surrogate, forbidden control and tab are encoded'
	);
	expect(
		condition := TOF_Core.Strings.Contains(stringToSearchIn := content^, stringToFind := 'END_OF_XML_DIAGNOSTIC'),
		message := 'Diagnostic suffix beyond 255 characters survives'
	);
	expect(
		condition := TOF_Core.Strings.Contains(stringToSearchIn := content^, stringToFind := 'time="1.250"'),
		message := 'JUnit duration uses decimal seconds'
	);
END_IF

checkXmlEncoding := TRUE;
END_METHOD

(*!
<summary>Repeats a nested run and checks configured and completed leaf counts, cleanup and escaped JUnit output.</summary>
<description>Configures owned fixtures through borrowed references without copying their state.
Returns TRUE when all observations for this scenario are complete.
</description>
*)
METHOD PRIVATE runAndCheck : BOOL
VAR
	content : POINTER TO STRING;
	probe : REFERENCE TO TestingProbe;
	multiCycleProbe : REFERENCE TO AssertionIsolationProbe;
END_VAR
IF NOT _Configured THEN
	expectDInt(expected := 5, actual := _Runner.FailureOuter.TestCount, message := 'Nested leaf count');
	expectDInt(expected := 0, actual := _Runner.Empty.TestCount, message := 'Empty group leaf count');
	expectDInt(expected := 1, actual := _Runner.Pass.TestCount, message := 'Single-cycle leaf count');
	expectDInt(expected := 1, actual := _Runner.Multi.TestCount, message := 'Multi-cycle leaf count');

	probe REF= _Runner.FailureOuter.Failures.SetupFailure;
	probe.ThrowBeforeTest := TRUE;
	probe REF= _Runner.FailureOuter.Failures.BodyFailure;
	probe.ThrowBody := TRUE;
	probe REF= _Runner.FailureOuter.Failures.TeardownFailure;
	probe.ThrowAfterTest := TRUE;
	probe REF= _Runner.FailureOuter.Failures.ComparisonFailure;
	probe.InvalidComparison := TRUE;
	probe REF= _Runner.FailureOuter.Failures.DiagnosticFailure;
	probe.DiagnosticFailure := TRUE;
	_Runner.Reporter := _Reporter;
	multiCycleProbe REF= _Runner.Multi;
	multiCycleProbe.Timeout := T#0S;
	_Configured := TRUE;
END_IF

_Runner.Execute(cleanupTaskMemory := FALSE);
_Calls := _Calls + 1;

IF NOT _Runner.IsFinished AND_THEN _Calls < 32 THEN
	RETURN;
END_IF

expect(condition := _Runner.IsFinished, message := 'The tree finishes within 32 scans');
expectDInt(expected := 2, actual := _Runner.PassedTests, message := 'Single and multi-cycle leaves pass');
expectDInt(expected := 5, actual := _Runner.FailedTests, message := 'Five distinct leaf failures');
expectDInt(expected := 7, actual := _Runner.TotalTests, message := 'Groups add no synthetic tests');
expectDInt(expected := 5, actual := _Runner.FailureOuter.TestCount, message := 'Leaf count survives a run');
expectUDInt(
	expected := 0,
	actual := _Runner.FailureOuter.Failures.SetupFailure.BodyCalls,
	message := 'Failed setup suppresses body'
);
expectUDInt(
	expected := 1,
	actual := _Runner.FailureOuter.Failures.SetupFailure.TeardownCalls,
	message := 'Failed setup still cleans up'
);
expectUDInt(
	expected := 1,
	actual := _Runner.FailureOuter.Failures.BodyFailure.TeardownCalls,
	message := 'Thrown body cleans up'
);
expectUDInt(
	expected := 1,
	actual := _Runner.FailureOuter.Failures.TeardownFailure.TeardownCalls,
	message := 'Thrown teardown is not retried'
);
expectUDInt(
	expected := 1,
	actual := _Runner.Pass.BodyCalls,
	message := 'Single-cycle body executes once per run'
);
expectUDInt(
	expected := 3,
	actual := _Runner.Multi.BodyCalls,
	message := 'Multi-cycle state survives three scans'
);
expectDInt(
	expected := 0,
	actual := _Runner.Empty.FailedCount,
	message := 'An empty group passes without tests'
);
expect(condition := _Reporter.IsReady, message := 'JUnit output is complete');
expect(
	condition := TOF_Core.WideStrings.Contains(stringToSearchIn := _Runner.FailureOuter.Failures.SetupFailure.FailureMessage,
		stringToFind := "BeforeTest: "),
	message := 'Preparation stage survives exception capture'
);
expect(
	condition := TOF_Core.WideStrings.Contains(stringToSearchIn := _Runner.FailureOuter.Failures.BodyFailure.FailureMessage,
		stringToFind := "Body failed"),
	message := 'Framework payload survives task cleanup'
);
expect(
	condition := TOF_Core.WideStrings.Contains(stringToSearchIn := _Runner.FailureOuter.Failures.BodyFailure.FailureMessage,
		stringToFind := "ExecuteTest"),
	message := 'Framework source survives task cleanup'
);
expect(
	condition := TOF_Core.WideStrings.Contains(stringToSearchIn := _Runner.FailureOuter.Failures.TeardownFailure.FailureMessage,
		stringToFind := "Teardown failed"),
	message := 'Teardown payload is copied'
);

content := _Reporter.ContentAddress;
expect(condition := content <> 0, message := 'Completed XML exposes a buffer');

IF content <> 0 THEN
	expect(
		condition := TOF_Core.Strings.Contains(
			stringToSearchIn := content^,
			stringToFind := 'Expected value &lt; '
		),
		message := 'An incompatible borrowed comparison remains an assertion failure'
	);
	expect(
		condition := TOF_Core.Strings.Contains(stringToSearchIn := content^, stringToFind := '&#1070;&amp;&lt;'),
		message := 'Cyrillic and XML markup are preserved'
	);
	expect(
		condition := TOF_Core.Strings.Contains(stringToSearchIn := content^, stringToFind := 'name=""'),
		message := 'Empty test name serializes safely'
	);
	expect(
		condition := TOF_Core.Strings.Contains(stringToSearchIn := content^, stringToFind := 'classname="Nested/Failures"'),
		message := 'The nested group path is preserved'
	);
END_IF

IF NOT _Repeated AND_THEN _Runner.IsFinished THEN
	_Repeated := TRUE;
	_Calls := 0;
	_Runner.Reset();
	RETURN;
END_IF

runAndCheck := TRUE;
END_METHOD

(*!
<summary>Borrows the initialized concrete class name.</summary>
*)
{attribute 'monitoring' := 'call'}
PROPERTY ClassName : REFERENCE TO STRING
GET
ClassName REF= _ClassName;
END_GET
END_PROPERTY

(*!
<summary>Borrows the project namespace name.</summary>
*)
{attribute 'monitoring' := 'call'}
PROPERTY NamespaceName : REFERENCE TO STRING
GET
NamespaceName REF= CurrentNamespace.Name;
END_GET
END_PROPERTY

END_FUNCTION_BLOCK

(* stored: Version 1.1.0.1
   POU TestRunnerContractTest: Id {fa92aa2f-994b-4ea4-8ec9-dcb12a01dbad}, SpecialFunc None
   Method Execute: Id {e31d9ffe-7b1b-45a2-9a00-a80f0b0e915e}
   Method expect: Id {9d28e443-da3c-4418-bcea-1b995d08f2ea}
   Method expectFalse: Id {8e44a3ee-f8e1-4ce0-93f5-068a46e2571a}
   Method expectDInt: Id {50b05224-dc7d-45b6-a273-dc7438b9c953}
   Method expectUDInt: Id {15c60658-7cd3-4324-92b4-c27644035f85}
   Method logResult: Id {221fc805-89ef-4d1b-bef5-27bda27c6307}
   Method assertCaughtExceptionType: Id {15ca4a6f-8e18-4c5c-a5c2-1bc97e01dba9}
   Method assertObjectMetadata: Id {b2db19e0-9754-403c-82ec-2e3c775ebec1}
   Method checkAssertionContracts: Id {d9e564a2-612e-4b45-b34a-fee9bbbe15b9}
   Method checkCaseIsolation: Id {515aeddf-ccd1-46f9-8790-e38279d4e123}
   Method checkContextObjects: Id {d30b1f3c-17b2-4908-91a0-da30356d6c6d}
   Method checkDeadline: Id {e519027d-6763-4eea-87bf-bb55734f0f09}
   Method checkDiagnostics: Id {b112f57d-7cbf-48a5-b2ae-60e53dfe141d}
   Method checkEmptyRun: Id {e4ed030a-bca3-4b47-b902-6f3f6606af4e}
   Method checkExceptionClasses: Id {c32f96d7-29ff-4026-aa6c-87146ca43581}
   Method checkAdsReporterSummary: Id {c2b70e83-8302-42c3-8b45-483cb8e41095}
   Method checkExternalRecovery: Id {c7b6aba0-ab1a-4823-b18b-979f2d38a5be}
   Method checkIndexedChildren: Id {ff86329b-fcb6-47e8-9300-27cf974a301e}
   Method checkPaths: Id {0d629b2f-c97c-49bb-a00e-9ed412fe9695}
   Method checkReporterAbort: Id {ff8cf1a3-fd79-4c4f-9137-e06eee3d3007}
   Method checkRunnerTopology: Id {0e7d627d-20a9-4651-8595-4eb23ecf183f}
   Method checkTopology: Id {e96454fa-d33d-44fe-a289-bf444e91ec4d}
   Method checkXmlEncoding: Id {a12404ad-44dd-4844-8d07-6492b26dc063}
   Method runAndCheck: Id {6e7eb7a7-8c88-4484-9a49-990753348b68}
   Property ClassName: Id {eb0a75ac-d210-47dd-990e-c97e2b015735}
   Get Get: Id {7c24322f-87c5-42ef-bb71-a244580d5210}
   Property NamespaceName: Id {1d0c31c3-44e2-4222-aa53-2cabfe5af769}
   Get Get: Id {70c6cd04-7621-4b43-9d4f-8c719b5bad9a} *)
